(* IEC 61131-3 sources: TetherPLC/compat/tc2 (part 4) *)

(* ---- tc2_modbussrv.st ---- *)
// Tc2_ModbusSrv Modbus client FBs (TwinCAT 3 PLC Library
// Tc2_ModbusSrv). Beckhoff-shaped wrappers over the builtin
// FB_Modbus, which drives the host "tplc-modbus" service
// (Modbus TCP and UDP, nonblocking, connect-per-transaction for
// TCP, one datagram per transaction for UDP).
// Differences from TwinCAT, documented in docs/plc/compat/README.md:
//   - POINTER TO BYTE payloads are ARRAY[0..255] OF BYTE buffers
//     (bounded; cbLength/cbSrcLength/cbDestLength still apply).
//   - sIPAddr is sHost (IPv4 dotted quad; no DNS).
//   - nErrId carries tplc-modbus transport codes, or the Modbus
//     exception code when the slave returns an exception response.
//   - Coil/register payloads are raw big-endian bytes; bit packing
//     for coil arrays is the caller's job, as in TwinCAT.
//   - the FB_MBUdp* wrappers below use the same ADU per UDP datagram
//     (MBAP+PDU); TwinCAT UDP encapsulation is assumed identical.
//   - the RTU library (Tc2_ModbusRTU) is not provided.
// Sources: docs/plc/plan/21-twincat-libraries.md §7 (TF6250).

FUNCTION_BLOCK FB_MBReadCoils
VAR_INPUT
    sHost : STRING[15];
    nTCPPort : UINT := 502;
    nUnitID : BYTE := 16#FF;
    nQuantity : WORD;
    nMBAddr : WORD;
    cbLength : UDINT;
    bExecute : BOOL;
    tTimeout : TIME;
END_VAR
VAR_OUTPUT
    bBusy : BOOL;
    bDone : BOOL;
    bError : BOOL;
    nErrId : UDINT;
    cbRead : UDINT;
    pData : ARRAY[0..255] OF BYTE;
END_VAR
VAR
    mb : FB_Modbus;
    i : UDINT;
END_VAR
    mb.FUNC := 1;
    mb.HOST := sHost;
    mb.PORT := nTCPPort;
    mb.UNIT := nUnitID;
    mb.TIMEOUT := tTimeout;
    mb.DATA[0] := UINT_TO_BYTE(nMBAddr / 256);
    mb.DATA[1] := UINT_TO_BYTE(nMBAddr MOD 256);
    mb.DATA[2] := UINT_TO_BYTE(nQuantity / 256);
    mb.DATA[3] := UINT_TO_BYTE(nQuantity MOD 256);
    mb.RLEN := 4;
    mb.EXEC := bExecute;
    mb();
    bBusy := mb.BUSY;
    bDone := mb.DONE;
    IF mb.DONE THEN
        i := 0;
        WHILE i < mb.DLEN AND i < 256 DO
            pData[i] := mb.DATA[i];
            i := i + 1;
        END_WHILE;
        cbRead := mb.DLEN;
    END_IF;
    nErrId := mb.ERRID;
    IF mb.RESULT = 1 THEN
        nErrId := 16#8000 + mb.EXC;
    END_IF;
    bError := (mb.ERRID <> 0) OR (mb.RESULT = 1);
END_FUNCTION_BLOCK

FUNCTION_BLOCK FB_MBReadInputs
VAR_INPUT
    sHost : STRING[15];
    nTCPPort : UINT := 502;
    nUnitID : BYTE := 16#FF;
    nQuantity : WORD;
    nMBAddr : WORD;
    cbLength : UDINT;
    bExecute : BOOL;
    tTimeout : TIME;
END_VAR
VAR_OUTPUT
    bBusy : BOOL;
    bDone : BOOL;
    bError : BOOL;
    nErrId : UDINT;
    cbRead : UDINT;
    pData : ARRAY[0..255] OF BYTE;
END_VAR
VAR
    mb : FB_Modbus;
    i : UDINT;
END_VAR
    mb.FUNC := 2;
    mb.HOST := sHost;
    mb.PORT := nTCPPort;
    mb.UNIT := nUnitID;
    mb.TIMEOUT := tTimeout;
    mb.DATA[0] := UINT_TO_BYTE(nMBAddr / 256);
    mb.DATA[1] := UINT_TO_BYTE(nMBAddr MOD 256);
    mb.DATA[2] := UINT_TO_BYTE(nQuantity / 256);
    mb.DATA[3] := UINT_TO_BYTE(nQuantity MOD 256);
    mb.RLEN := 4;
    mb.EXEC := bExecute;
    mb();
    bBusy := mb.BUSY;
    bDone := mb.DONE;
    IF mb.DONE THEN
        i := 0;
        WHILE i < mb.DLEN AND i < 256 DO
            pData[i] := mb.DATA[i];
            i := i + 1;
        END_WHILE;
        cbRead := mb.DLEN;
    END_IF;
    nErrId := mb.ERRID;
    IF mb.RESULT = 1 THEN
        nErrId := 16#8000 + mb.EXC;
    END_IF;
    bError := (mb.ERRID <> 0) OR (mb.RESULT = 1);
END_FUNCTION_BLOCK

FUNCTION_BLOCK FB_MBReadRegs
VAR_INPUT
    sHost : STRING[15];
    nTCPPort : UINT := 502;
    nUnitID : BYTE := 16#FF;
    nQuantity : WORD;
    nMBAddr : WORD;
    cbLength : UDINT;
    bExecute : BOOL;
    tTimeout : TIME;
END_VAR
VAR_OUTPUT
    bBusy : BOOL;
    bDone : BOOL;
    bError : BOOL;
    nErrId : UDINT;
    cbRead : UDINT;
    pData : ARRAY[0..255] OF BYTE;
END_VAR
VAR
    mb : FB_Modbus;
    i : UDINT;
END_VAR
    mb.FUNC := 3;
    mb.HOST := sHost;
    mb.PORT := nTCPPort;
    mb.UNIT := nUnitID;
    mb.TIMEOUT := tTimeout;
    mb.DATA[0] := UINT_TO_BYTE(nMBAddr / 256);
    mb.DATA[1] := UINT_TO_BYTE(nMBAddr MOD 256);
    mb.DATA[2] := UINT_TO_BYTE(nQuantity / 256);
    mb.DATA[3] := UINT_TO_BYTE(nQuantity MOD 256);
    mb.RLEN := 4;
    mb.EXEC := bExecute;
    mb();
    bBusy := mb.BUSY;
    bDone := mb.DONE;
    IF mb.DONE THEN
        i := 0;
        WHILE i < mb.DLEN AND i < 256 DO
            pData[i] := mb.DATA[i];
            i := i + 1;
        END_WHILE;
        cbRead := mb.DLEN;
    END_IF;
    nErrId := mb.ERRID;
    IF mb.RESULT = 1 THEN
        nErrId := 16#8000 + mb.EXC;
    END_IF;
    bError := (mb.ERRID <> 0) OR (mb.RESULT = 1);
END_FUNCTION_BLOCK

FUNCTION_BLOCK FB_MBReadInputRegs
VAR_INPUT
    sHost : STRING[15];
    nTCPPort : UINT := 502;
    nUnitID : BYTE := 16#FF;
    nQuantity : WORD;
    nMBAddr : WORD;
    cbLength : UDINT;
    bExecute : BOOL;
    tTimeout : TIME;
END_VAR
VAR_OUTPUT
    bBusy : BOOL;
    bDone : BOOL;
    bError : BOOL;
    nErrId : UDINT;
    cbRead : UDINT;
    pData : ARRAY[0..255] OF BYTE;
END_VAR
VAR
    mb : FB_Modbus;
    i : UDINT;
END_VAR
    mb.FUNC := 4;
    mb.HOST := sHost;
    mb.PORT := nTCPPort;
    mb.UNIT := nUnitID;
    mb.TIMEOUT := tTimeout;
    mb.DATA[0] := UINT_TO_BYTE(nMBAddr / 256);
    mb.DATA[1] := UINT_TO_BYTE(nMBAddr MOD 256);
    mb.DATA[2] := UINT_TO_BYTE(nQuantity / 256);
    mb.DATA[3] := UINT_TO_BYTE(nQuantity MOD 256);
    mb.RLEN := 4;
    mb.EXEC := bExecute;
    mb();
    bBusy := mb.BUSY;
    bDone := mb.DONE;
    IF mb.DONE THEN
        i := 0;
        WHILE i < mb.DLEN AND i < 256 DO
            pData[i] := mb.DATA[i];
            i := i + 1;
        END_WHILE;
        cbRead := mb.DLEN;
    END_IF;
    nErrId := mb.ERRID;
    IF mb.RESULT = 1 THEN
        nErrId := 16#8000 + mb.EXC;
    END_IF;
    bError := (mb.ERRID <> 0) OR (mb.RESULT = 1);
END_FUNCTION_BLOCK

FUNCTION_BLOCK FB_MBWriteSingleCoil
VAR_INPUT
    sHost : STRING[15];
    nTCPPort : UINT := 502;
    nUnitID : BYTE := 16#FF;
    nMBAddr : WORD;
    nValue : WORD;
    bExecute : BOOL;
    tTimeout : TIME;
END_VAR
VAR_OUTPUT
    bBusy : BOOL;
    bDone : BOOL;
    bError : BOOL;
    nErrId : UDINT;
    cbRead : UDINT;
END_VAR
VAR
    mb : FB_Modbus;
END_VAR
    mb.FUNC := 5;
    mb.HOST := sHost;
    mb.PORT := nTCPPort;
    mb.UNIT := nUnitID;
    mb.TIMEOUT := tTimeout;
    mb.DATA[0] := UINT_TO_BYTE(nMBAddr / 256);
    mb.DATA[1] := UINT_TO_BYTE(nMBAddr MOD 256);
    mb.DATA[2] := UINT_TO_BYTE(nValue / 256);
    mb.DATA[3] := UINT_TO_BYTE(nValue MOD 256);
    mb.RLEN := 4;
    mb.EXEC := bExecute;
    mb();
    bBusy := mb.BUSY;
    bDone := mb.DONE;
    cbRead := 0;
    nErrId := mb.ERRID;
    IF mb.RESULT = 1 THEN
        nErrId := 16#8000 + mb.EXC;
    END_IF;
    bError := (mb.ERRID <> 0) OR (mb.RESULT = 1);
END_FUNCTION_BLOCK

FUNCTION_BLOCK FB_MBWriteSingleReg
VAR_INPUT
    sHost : STRING[15];
    nTCPPort : UINT := 502;
    nUnitID : BYTE := 16#FF;
    nMBAddr : WORD;
    nValue : WORD;
    bExecute : BOOL;
    tTimeout : TIME;
END_VAR
VAR_OUTPUT
    bBusy : BOOL;
    bDone : BOOL;
    bError : BOOL;
    nErrId : UDINT;
    cbRead : UDINT;
END_VAR
VAR
    mb : FB_Modbus;
END_VAR
    mb.FUNC := 6;
    mb.HOST := sHost;
    mb.PORT := nTCPPort;
    mb.UNIT := nUnitID;
    mb.TIMEOUT := tTimeout;
    mb.DATA[0] := UINT_TO_BYTE(nMBAddr / 256);
    mb.DATA[1] := UINT_TO_BYTE(nMBAddr MOD 256);
    mb.DATA[2] := UINT_TO_BYTE(nValue / 256);
    mb.DATA[3] := UINT_TO_BYTE(nValue MOD 256);
    mb.RLEN := 4;
    mb.EXEC := bExecute;
    mb();
    bBusy := mb.BUSY;
    bDone := mb.DONE;
    cbRead := 0;
    nErrId := mb.ERRID;
    IF mb.RESULT = 1 THEN
        nErrId := 16#8000 + mb.EXC;
    END_IF;
    bError := (mb.ERRID <> 0) OR (mb.RESULT = 1);
END_FUNCTION_BLOCK

FUNCTION_BLOCK FB_MBWriteCoils
VAR_INPUT
    sHost : STRING[15];
    nTCPPort : UINT := 502;
    nUnitID : BYTE := 16#FF;
    nQuantity : WORD;
    nMBAddr : WORD;
    cbLength : UDINT;
    pSrcData : ARRAY[0..255] OF BYTE;
    bExecute : BOOL;
    tTimeout : TIME;
END_VAR
VAR_OUTPUT
    bBusy : BOOL;
    bDone : BOOL;
    bError : BOOL;
    nErrId : UDINT;
    cbRead : UDINT;
END_VAR
VAR
    mb : FB_Modbus;
    i : UDINT;
    n : UDINT;
END_VAR
    mb.FUNC := 15;
    mb.HOST := sHost;
    mb.PORT := nTCPPort;
    mb.UNIT := nUnitID;
    mb.TIMEOUT := tTimeout;
    mb.DATA[0] := UINT_TO_BYTE(nMBAddr / 256);
    mb.DATA[1] := UINT_TO_BYTE(nMBAddr MOD 256);
    mb.DATA[2] := UINT_TO_BYTE(nQuantity / 256);
    mb.DATA[3] := UINT_TO_BYTE(nQuantity MOD 256);
    n := cbLength;
    IF n > 246 THEN
        n := 246;
    END_IF;
    mb.DATA[4] := UDINT_TO_BYTE(n);
    i := 0;
    WHILE i < n DO
        mb.DATA[5 + i] := pSrcData[i];
        i := i + 1;
    END_WHILE;
    mb.RLEN := 5 + n;
    mb.EXEC := bExecute;
    mb();
    bBusy := mb.BUSY;
    bDone := mb.DONE;
    cbRead := 0;
    nErrId := mb.ERRID;
    IF mb.RESULT = 1 THEN
        nErrId := 16#8000 + mb.EXC;
    END_IF;
    bError := (mb.ERRID <> 0) OR (mb.RESULT = 1);
END_FUNCTION_BLOCK

FUNCTION_BLOCK FB_MBWriteRegs
VAR_INPUT
    sHost : STRING[15];
    nTCPPort : UINT := 502;
    nUnitID : BYTE := 16#FF;
    nQuantity : WORD;
    nMBAddr : WORD;
    cbLength : UDINT;
    pSrcData : ARRAY[0..255] OF BYTE;
    bExecute : BOOL;
    tTimeout : TIME;
END_VAR
VAR_OUTPUT
    bBusy : BOOL;
    bDone : BOOL;
    bError : BOOL;
    nErrId : UDINT;
    cbRead : UDINT;
END_VAR
VAR
    mb : FB_Modbus;
    i : UDINT;
    n : UDINT;
END_VAR
    mb.FUNC := 16;
    mb.HOST := sHost;
    mb.PORT := nTCPPort;
    mb.UNIT := nUnitID;
    mb.TIMEOUT := tTimeout;
    mb.DATA[0] := UINT_TO_BYTE(nMBAddr / 256);
    mb.DATA[1] := UINT_TO_BYTE(nMBAddr MOD 256);
    mb.DATA[2] := UINT_TO_BYTE(nQuantity / 256);
    mb.DATA[3] := UINT_TO_BYTE(nQuantity MOD 256);
    n := cbLength;
    IF n > 246 THEN
        n := 246;
    END_IF;
    mb.DATA[4] := UDINT_TO_BYTE(n);
    i := 0;
    WHILE i < n DO
        mb.DATA[5 + i] := pSrcData[i];
        i := i + 1;
    END_WHILE;
    mb.RLEN := 5 + n;
    mb.EXEC := bExecute;
    mb();
    bBusy := mb.BUSY;
    bDone := mb.DONE;
    cbRead := 0;
    nErrId := mb.ERRID;
    IF mb.RESULT = 1 THEN
        nErrId := 16#8000 + mb.EXC;
    END_IF;
    bError := (mb.ERRID <> 0) OR (mb.RESULT = 1);
END_FUNCTION_BLOCK

FUNCTION_BLOCK FB_MBReadWriteRegs
VAR_INPUT
    sHost : STRING[15];
    nTCPPort : UINT := 502;
    nUnitID : BYTE := 16#FF;
    nReadQuantity : WORD;
    nMBReadAddr : WORD;
    nWriteQuantity : WORD;
    nMBWriteAddr : WORD;
    cbDestLength : UDINT;
    cbSrcLength : UDINT;
    pSrcData : ARRAY[0..255] OF BYTE;
    bExecute : BOOL;
    tTimeout : TIME;
END_VAR
VAR_OUTPUT
    bBusy : BOOL;
    bDone : BOOL;
    bError : BOOL;
    nErrId : UDINT;
    cbRead : UDINT;
    pDestData : ARRAY[0..255] OF BYTE;
END_VAR
VAR
    mb : FB_Modbus;
    i : UDINT;
    n : UDINT;
END_VAR
    mb.FUNC := 23;
    mb.HOST := sHost;
    mb.PORT := nTCPPort;
    mb.UNIT := nUnitID;
    mb.TIMEOUT := tTimeout;
    mb.DATA[0] := UINT_TO_BYTE(nMBReadAddr / 256);
    mb.DATA[1] := UINT_TO_BYTE(nMBReadAddr MOD 256);
    mb.DATA[2] := UINT_TO_BYTE(nReadQuantity / 256);
    mb.DATA[3] := UINT_TO_BYTE(nReadQuantity MOD 256);
    mb.DATA[4] := UINT_TO_BYTE(nMBWriteAddr / 256);
    mb.DATA[5] := UINT_TO_BYTE(nMBWriteAddr MOD 256);
    mb.DATA[6] := UINT_TO_BYTE(nWriteQuantity / 256);
    mb.DATA[7] := UINT_TO_BYTE(nWriteQuantity MOD 256);
    n := cbSrcLength;
    IF n > 242 THEN
        n := 242;
    END_IF;
    mb.DATA[8] := UDINT_TO_BYTE(n);
    i := 0;
    WHILE i < n DO
        mb.DATA[9 + i] := pSrcData[i];
        i := i + 1;
    END_WHILE;
    mb.RLEN := 9 + n;
    mb.EXEC := bExecute;
    mb();
    bBusy := mb.BUSY;
    bDone := mb.DONE;
    IF mb.DONE THEN
        i := 0;
        WHILE i < mb.DLEN AND i < 256 DO
            pDestData[i] := mb.DATA[i];
            i := i + 1;
        END_WHILE;
        cbRead := mb.DLEN;
    END_IF;
    nErrId := mb.ERRID;
    IF mb.RESULT = 1 THEN
        nErrId := 16#8000 + mb.EXC;
    END_IF;
    bError := (mb.ERRID <> 0) OR (mb.RESULT = 1);
END_FUNCTION_BLOCK

FUNCTION_BLOCK FB_MBDiagnose
VAR_INPUT
    sHost : STRING[15];
    nTCPPort : UINT := 502;
    nUnitID : BYTE := 16#FF;
    nWriteData : WORD;
    bExecute : BOOL;
    tTimeout : TIME;
END_VAR
VAR_OUTPUT
    bBusy : BOOL;
    bDone : BOOL;
    bError : BOOL;
    nErrId : UDINT;
    cbRead : UDINT;
    pData : ARRAY[0..255] OF BYTE;
END_VAR
VAR
    mb : FB_Modbus;
    i : UDINT;
END_VAR
    mb.FUNC := 8;
    mb.HOST := sHost;
    mb.PORT := nTCPPort;
    mb.UNIT := nUnitID;
    mb.TIMEOUT := tTimeout;
    mb.DATA[0] := UINT_TO_BYTE(nWriteData / 256);
    mb.DATA[1] := UINT_TO_BYTE(nWriteData MOD 256);
    mb.RLEN := 2;
    mb.EXEC := bExecute;
    mb();
    bBusy := mb.BUSY;
    bDone := mb.DONE;
    IF mb.DONE THEN
        i := 0;
        WHILE i < mb.DLEN AND i < 256 DO
            pData[i] := mb.DATA[i];
            i := i + 1;
        END_WHILE;
        cbRead := mb.DLEN;
    END_IF;
    nErrId := mb.ERRID;
    IF mb.RESULT = 1 THEN
        nErrId := 16#8000 + mb.EXC;
    END_IF;
    bError := (mb.ERRID <> 0) OR (mb.RESULT = 1);
END_FUNCTION_BLOCK
FUNCTION_BLOCK FB_MBUdpReadCoils
VAR_INPUT
    sHost : STRING[15];
    nTCPPort : UINT := 502;
    nUnitID : BYTE := 16#FF;
    nQuantity : WORD;
    nMBAddr : WORD;
    cbLength : UDINT;
    bExecute : BOOL;
    tTimeout : TIME;
END_VAR
VAR_OUTPUT
    bBusy : BOOL;
    bDone : BOOL;
    bError : BOOL;
    nErrId : UDINT;
    cbRead : UDINT;
    pData : ARRAY[0..255] OF BYTE;
END_VAR
VAR
    mb : FB_Modbus;
    i : UDINT;
END_VAR
    mb.FUNC := 1;
    mb.HOST := sHost;
    mb.PORT := nTCPPort;
    mb.UNIT := nUnitID;
    mb.TIMEOUT := tTimeout;
    mb.DATA[0] := UINT_TO_BYTE(nMBAddr / 256);
    mb.DATA[1] := UINT_TO_BYTE(nMBAddr MOD 256);
    mb.DATA[2] := UINT_TO_BYTE(nQuantity / 256);
    mb.DATA[3] := UINT_TO_BYTE(nQuantity MOD 256);
    mb.RLEN := 4;
    mb.UDP := TRUE;
    mb.EXEC := bExecute;
    mb();
    bBusy := mb.BUSY;
    bDone := mb.DONE;
    IF mb.DONE THEN
        i := 0;
        WHILE i < mb.DLEN AND i < 256 DO
            pData[i] := mb.DATA[i];
            i := i + 1;
        END_WHILE;
        cbRead := mb.DLEN;
    END_IF;
    nErrId := mb.ERRID;
    IF mb.RESULT = 1 THEN
        nErrId := 16#8000 + mb.EXC;
    END_IF;
    bError := (mb.ERRID <> 0) OR (mb.RESULT = 1);
END_FUNCTION_BLOCK

FUNCTION_BLOCK FB_MBUdpReadInputs
VAR_INPUT
    sHost : STRING[15];
    nTCPPort : UINT := 502;
    nUnitID : BYTE := 16#FF;
    nQuantity : WORD;
    nMBAddr : WORD;
    cbLength : UDINT;
    bExecute : BOOL;
    tTimeout : TIME;
END_VAR
VAR_OUTPUT
    bBusy : BOOL;
    bDone : BOOL;
    bError : BOOL;
    nErrId : UDINT;
    cbRead : UDINT;
    pData : ARRAY[0..255] OF BYTE;
END_VAR
VAR
    mb : FB_Modbus;
    i : UDINT;
END_VAR
    mb.FUNC := 2;
    mb.HOST := sHost;
    mb.PORT := nTCPPort;
    mb.UNIT := nUnitID;
    mb.TIMEOUT := tTimeout;
    mb.DATA[0] := UINT_TO_BYTE(nMBAddr / 256);
    mb.DATA[1] := UINT_TO_BYTE(nMBAddr MOD 256);
    mb.DATA[2] := UINT_TO_BYTE(nQuantity / 256);
    mb.DATA[3] := UINT_TO_BYTE(nQuantity MOD 256);
    mb.RLEN := 4;
    mb.UDP := TRUE;
    mb.EXEC := bExecute;
    mb();
    bBusy := mb.BUSY;
    bDone := mb.DONE;
    IF mb.DONE THEN
        i := 0;
        WHILE i < mb.DLEN AND i < 256 DO
            pData[i] := mb.DATA[i];
            i := i + 1;
        END_WHILE;
        cbRead := mb.DLEN;
    END_IF;
    nErrId := mb.ERRID;
    IF mb.RESULT = 1 THEN
        nErrId := 16#8000 + mb.EXC;
    END_IF;
    bError := (mb.ERRID <> 0) OR (mb.RESULT = 1);
END_FUNCTION_BLOCK

FUNCTION_BLOCK FB_MBUdpReadRegs
VAR_INPUT
    sHost : STRING[15];
    nTCPPort : UINT := 502;
    nUnitID : BYTE := 16#FF;
    nQuantity : WORD;
    nMBAddr : WORD;
    cbLength : UDINT;
    bExecute : BOOL;
    tTimeout : TIME;
END_VAR
VAR_OUTPUT
    bBusy : BOOL;
    bDone : BOOL;
    bError : BOOL;
    nErrId : UDINT;
    cbRead : UDINT;
    pData : ARRAY[0..255] OF BYTE;
END_VAR
VAR
    mb : FB_Modbus;
    i : UDINT;
END_VAR
    mb.FUNC := 3;
    mb.HOST := sHost;
    mb.PORT := nTCPPort;
    mb.UNIT := nUnitID;
    mb.TIMEOUT := tTimeout;
    mb.DATA[0] := UINT_TO_BYTE(nMBAddr / 256);
    mb.DATA[1] := UINT_TO_BYTE(nMBAddr MOD 256);
    mb.DATA[2] := UINT_TO_BYTE(nQuantity / 256);
    mb.DATA[3] := UINT_TO_BYTE(nQuantity MOD 256);
    mb.RLEN := 4;
    mb.UDP := TRUE;
    mb.EXEC := bExecute;
    mb();
    bBusy := mb.BUSY;
    bDone := mb.DONE;
    IF mb.DONE THEN
        i := 0;
        WHILE i < mb.DLEN AND i < 256 DO
            pData[i] := mb.DATA[i];
            i := i + 1;
        END_WHILE;
        cbRead := mb.DLEN;
    END_IF;
    nErrId := mb.ERRID;
    IF mb.RESULT = 1 THEN
        nErrId := 16#8000 + mb.EXC;
    END_IF;
    bError := (mb.ERRID <> 0) OR (mb.RESULT = 1);
END_FUNCTION_BLOCK

FUNCTION_BLOCK FB_MBUdpReadInputRegs
VAR_INPUT
    sHost : STRING[15];
    nTCPPort : UINT := 502;
    nUnitID : BYTE := 16#FF;
    nQuantity : WORD;
    nMBAddr : WORD;
    cbLength : UDINT;
    bExecute : BOOL;
    tTimeout : TIME;
END_VAR
VAR_OUTPUT
    bBusy : BOOL;
    bDone : BOOL;
    bError : BOOL;
    nErrId : UDINT;
    cbRead : UDINT;
    pData : ARRAY[0..255] OF BYTE;
END_VAR
VAR
    mb : FB_Modbus;
    i : UDINT;
END_VAR
    mb.FUNC := 4;
    mb.HOST := sHost;
    mb.PORT := nTCPPort;
    mb.UNIT := nUnitID;
    mb.TIMEOUT := tTimeout;
    mb.DATA[0] := UINT_TO_BYTE(nMBAddr / 256);
    mb.DATA[1] := UINT_TO_BYTE(nMBAddr MOD 256);
    mb.DATA[2] := UINT_TO_BYTE(nQuantity / 256);
    mb.DATA[3] := UINT_TO_BYTE(nQuantity MOD 256);
    mb.RLEN := 4;
    mb.UDP := TRUE;
    mb.EXEC := bExecute;
    mb();
    bBusy := mb.BUSY;
    bDone := mb.DONE;
    IF mb.DONE THEN
        i := 0;
        WHILE i < mb.DLEN AND i < 256 DO
            pData[i] := mb.DATA[i];
            i := i + 1;
        END_WHILE;
        cbRead := mb.DLEN;
    END_IF;
    nErrId := mb.ERRID;
    IF mb.RESULT = 1 THEN
        nErrId := 16#8000 + mb.EXC;
    END_IF;
    bError := (mb.ERRID <> 0) OR (mb.RESULT = 1);
END_FUNCTION_BLOCK

FUNCTION_BLOCK FB_MBUdpWriteSingleCoil
VAR_INPUT
    sHost : STRING[15];
    nTCPPort : UINT := 502;
    nUnitID : BYTE := 16#FF;
    nMBAddr : WORD;
    nValue : WORD;
    bExecute : BOOL;
    tTimeout : TIME;
END_VAR
VAR_OUTPUT
    bBusy : BOOL;
    bDone : BOOL;
    bError : BOOL;
    nErrId : UDINT;
    cbRead : UDINT;
END_VAR
VAR
    mb : FB_Modbus;
END_VAR
    mb.FUNC := 5;
    mb.HOST := sHost;
    mb.PORT := nTCPPort;
    mb.UNIT := nUnitID;
    mb.TIMEOUT := tTimeout;
    mb.DATA[0] := UINT_TO_BYTE(nMBAddr / 256);
    mb.DATA[1] := UINT_TO_BYTE(nMBAddr MOD 256);
    mb.DATA[2] := UINT_TO_BYTE(nValue / 256);
    mb.DATA[3] := UINT_TO_BYTE(nValue MOD 256);
    mb.RLEN := 4;
    mb.UDP := TRUE;
    mb.EXEC := bExecute;
    mb();
    bBusy := mb.BUSY;
    bDone := mb.DONE;
    cbRead := 0;
    nErrId := mb.ERRID;
    IF mb.RESULT = 1 THEN
        nErrId := 16#8000 + mb.EXC;
    END_IF;
    bError := (mb.ERRID <> 0) OR (mb.RESULT = 1);
END_FUNCTION_BLOCK

FUNCTION_BLOCK FB_MBUdpWriteSingleReg
VAR_INPUT
    sHost : STRING[15];
    nTCPPort : UINT := 502;
    nUnitID : BYTE := 16#FF;
    nMBAddr : WORD;
    nValue : WORD;
    bExecute : BOOL;
    tTimeout : TIME;
END_VAR
VAR_OUTPUT
    bBusy : BOOL;
    bDone : BOOL;
    bError : BOOL;
    nErrId : UDINT;
    cbRead : UDINT;
END_VAR
VAR
    mb : FB_Modbus;
END_VAR
    mb.FUNC := 6;
    mb.HOST := sHost;
    mb.PORT := nTCPPort;
    mb.UNIT := nUnitID;
    mb.TIMEOUT := tTimeout;
    mb.DATA[0] := UINT_TO_BYTE(nMBAddr / 256);
    mb.DATA[1] := UINT_TO_BYTE(nMBAddr MOD 256);
    mb.DATA[2] := UINT_TO_BYTE(nValue / 256);
    mb.DATA[3] := UINT_TO_BYTE(nValue MOD 256);
    mb.RLEN := 4;
    mb.UDP := TRUE;
    mb.EXEC := bExecute;
    mb();
    bBusy := mb.BUSY;
    bDone := mb.DONE;
    cbRead := 0;
    nErrId := mb.ERRID;
    IF mb.RESULT = 1 THEN
        nErrId := 16#8000 + mb.EXC;
    END_IF;
    bError := (mb.ERRID <> 0) OR (mb.RESULT = 1);
END_FUNCTION_BLOCK

FUNCTION_BLOCK FB_MBUdpWriteCoils
VAR_INPUT
    sHost : STRING[15];
    nTCPPort : UINT := 502;
    nUnitID : BYTE := 16#FF;
    nQuantity : WORD;
    nMBAddr : WORD;
    cbLength : UDINT;
    pSrcData : ARRAY[0..255] OF BYTE;
    bExecute : BOOL;
    tTimeout : TIME;
END_VAR
VAR_OUTPUT
    bBusy : BOOL;
    bDone : BOOL;
    bError : BOOL;
    nErrId : UDINT;
    cbRead : UDINT;
END_VAR
VAR
    mb : FB_Modbus;
    i : UDINT;
    n : UDINT;
END_VAR
    mb.FUNC := 15;
    mb.HOST := sHost;
    mb.PORT := nTCPPort;
    mb.UNIT := nUnitID;
    mb.TIMEOUT := tTimeout;
    mb.DATA[0] := UINT_TO_BYTE(nMBAddr / 256);
    mb.DATA[1] := UINT_TO_BYTE(nMBAddr MOD 256);
    mb.DATA[2] := UINT_TO_BYTE(nQuantity / 256);
    mb.DATA[3] := UINT_TO_BYTE(nQuantity MOD 256);
    n := cbLength;
    IF n > 246 THEN
        n := 246;
    END_IF;
    mb.DATA[4] := UDINT_TO_BYTE(n);
    i := 0;
    WHILE i < n DO
        mb.DATA[5 + i] := pSrcData[i];
        i := i + 1;
    END_WHILE;
    mb.RLEN := 5 + n;
    mb.UDP := TRUE;
    mb.EXEC := bExecute;
    mb();
    bBusy := mb.BUSY;
    bDone := mb.DONE;
    cbRead := 0;
    nErrId := mb.ERRID;
    IF mb.RESULT = 1 THEN
        nErrId := 16#8000 + mb.EXC;
    END_IF;
    bError := (mb.ERRID <> 0) OR (mb.RESULT = 1);
END_FUNCTION_BLOCK

FUNCTION_BLOCK FB_MBUdpWriteRegs
VAR_INPUT
    sHost : STRING[15];
    nTCPPort : UINT := 502;
    nUnitID : BYTE := 16#FF;
    nQuantity : WORD;
    nMBAddr : WORD;
    cbLength : UDINT;
    pSrcData : ARRAY[0..255] OF BYTE;
    bExecute : BOOL;
    tTimeout : TIME;
END_VAR
VAR_OUTPUT
    bBusy : BOOL;
    bDone : BOOL;
    bError : BOOL;
    nErrId : UDINT;
    cbRead : UDINT;
END_VAR
VAR
    mb : FB_Modbus;
    i : UDINT;
    n : UDINT;
END_VAR
    mb.FUNC := 16;
    mb.HOST := sHost;
    mb.PORT := nTCPPort;
    mb.UNIT := nUnitID;
    mb.TIMEOUT := tTimeout;
    mb.DATA[0] := UINT_TO_BYTE(nMBAddr / 256);
    mb.DATA[1] := UINT_TO_BYTE(nMBAddr MOD 256);
    mb.DATA[2] := UINT_TO_BYTE(nQuantity / 256);
    mb.DATA[3] := UINT_TO_BYTE(nQuantity MOD 256);
    n := cbLength;
    IF n > 246 THEN
        n := 246;
    END_IF;
    mb.DATA[4] := UDINT_TO_BYTE(n);
    i := 0;
    WHILE i < n DO
        mb.DATA[5 + i] := pSrcData[i];
        i := i + 1;
    END_WHILE;
    mb.RLEN := 5 + n;
    mb.UDP := TRUE;
    mb.EXEC := bExecute;
    mb();
    bBusy := mb.BUSY;
    bDone := mb.DONE;
    cbRead := 0;
    nErrId := mb.ERRID;
    IF mb.RESULT = 1 THEN
        nErrId := 16#8000 + mb.EXC;
    END_IF;
    bError := (mb.ERRID <> 0) OR (mb.RESULT = 1);
END_FUNCTION_BLOCK

FUNCTION_BLOCK FB_MBUdpReadWriteRegs
VAR_INPUT
    sHost : STRING[15];
    nTCPPort : UINT := 502;
    nUnitID : BYTE := 16#FF;
    nReadQuantity : WORD;
    nMBReadAddr : WORD;
    nWriteQuantity : WORD;
    nMBWriteAddr : WORD;
    cbDestLength : UDINT;
    cbSrcLength : UDINT;
    pSrcData : ARRAY[0..255] OF BYTE;
    bExecute : BOOL;
    tTimeout : TIME;
END_VAR
VAR_OUTPUT
    bBusy : BOOL;
    bDone : BOOL;
    bError : BOOL;
    nErrId : UDINT;
    cbRead : UDINT;
    pDestData : ARRAY[0..255] OF BYTE;
END_VAR
VAR
    mb : FB_Modbus;
    i : UDINT;
    n : UDINT;
END_VAR
    mb.FUNC := 23;
    mb.HOST := sHost;
    mb.PORT := nTCPPort;
    mb.UNIT := nUnitID;
    mb.TIMEOUT := tTimeout;
    mb.DATA[0] := UINT_TO_BYTE(nMBReadAddr / 256);
    mb.DATA[1] := UINT_TO_BYTE(nMBReadAddr MOD 256);
    mb.DATA[2] := UINT_TO_BYTE(nReadQuantity / 256);
    mb.DATA[3] := UINT_TO_BYTE(nReadQuantity MOD 256);
    mb.DATA[4] := UINT_TO_BYTE(nMBWriteAddr / 256);
    mb.DATA[5] := UINT_TO_BYTE(nMBWriteAddr MOD 256);
    mb.DATA[6] := UINT_TO_BYTE(nWriteQuantity / 256);
    mb.DATA[7] := UINT_TO_BYTE(nWriteQuantity MOD 256);
    n := cbSrcLength;
    IF n > 242 THEN
        n := 242;
    END_IF;
    mb.DATA[8] := UDINT_TO_BYTE(n);
    i := 0;
    WHILE i < n DO
        mb.DATA[9 + i] := pSrcData[i];
        i := i + 1;
    END_WHILE;
    mb.RLEN := 9 + n;
    mb.UDP := TRUE;
    mb.EXEC := bExecute;
    mb();
    bBusy := mb.BUSY;
    bDone := mb.DONE;
    IF mb.DONE THEN
        i := 0;
        WHILE i < mb.DLEN AND i < 256 DO
            pDestData[i] := mb.DATA[i];
            i := i + 1;
        END_WHILE;
        cbRead := mb.DLEN;
    END_IF;
    nErrId := mb.ERRID;
    IF mb.RESULT = 1 THEN
        nErrId := 16#8000 + mb.EXC;
    END_IF;
    bError := (mb.ERRID <> 0) OR (mb.RESULT = 1);
END_FUNCTION_BLOCK

FUNCTION_BLOCK FB_MBUdpDiagnose
VAR_INPUT
    sHost : STRING[15];
    nTCPPort : UINT := 502;
    nUnitID : BYTE := 16#FF;
    nWriteData : WORD;
    bExecute : BOOL;
    tTimeout : TIME;
END_VAR
VAR_OUTPUT
    bBusy : BOOL;
    bDone : BOOL;
    bError : BOOL;
    nErrId : UDINT;
    cbRead : UDINT;
    pData : ARRAY[0..255] OF BYTE;
END_VAR
VAR
    mb : FB_Modbus;
    i : UDINT;
END_VAR
    mb.FUNC := 8;
    mb.HOST := sHost;
    mb.PORT := nTCPPort;
    mb.UNIT := nUnitID;
    mb.TIMEOUT := tTimeout;
    mb.DATA[0] := UINT_TO_BYTE(nWriteData / 256);
    mb.DATA[1] := UINT_TO_BYTE(nWriteData MOD 256);
    mb.RLEN := 2;
    mb.UDP := TRUE;
    mb.EXEC := bExecute;
    mb();
    bBusy := mb.BUSY;
    bDone := mb.DONE;
    IF mb.DONE THEN
        i := 0;
        WHILE i < mb.DLEN AND i < 256 DO
            pData[i] := mb.DATA[i];
            i := i + 1;
        END_WHILE;
        cbRead := mb.DLEN;
    END_IF;
    nErrId := mb.ERRID;
    IF mb.RESULT = 1 THEN
        nErrId := 16#8000 + mb.EXC;
    END_IF;
    bError := (mb.ERRID <> 0) OR (mb.RESULT = 1);
END_FUNCTION_BLOCK

(* ---- tc2_mpbus.st ---- *)
// tc2_mpbus.st — Tc2_MPBus surface (TwinCAT_3_PLC_Lib_Tc2_
// MPBus_EN): Belimo MP-Bus master over an opt-in serial adapter
// (9600 8N1, e.g. a USB MP-Bus gateway presenting a tty — the
// KL6771 terminal's process image is not modeled).  Wire
// format: [DA][CMD][LEN][data][CHK8-xor] request/response
// frames; the transact op sends and captures the reply.
//
// Differences (docs/plc/compat/README.md):
//   - The KL6771 bus-terminal process image is replaced by a
//     serial MP-Bus adapter — the function blocks take a PortHdl
//     from FB_MpbusOpen instead of terminal IO arrays.
//   - The full Belimo device-profile command matrix (Energy
//     Valve, CMV, addressing wizards) is simplified to raw
//     command ids; profile semantics are a documented gap.

// ---- FB_MpbusOpen: open the serial MP-Bus adapter ----
FUNCTION_BLOCK FB_MpbusOpen
VAR_INPUT
    Execute : BOOL;
    Path : STRING;
END_VAR
VAR_OUTPUT
    Done : BOOL;
    Error : BOOL;
    ErrorID : UDINT;
    PortHdl : UDINT;
END_VAR
VAR
    ch : FB_Mpbus;
END_VAR
    Done := FALSE;
    Error := FALSE;
    ErrorID := 0;
    IF Execute THEN
        ch.OP := 1;
        ch.PATH := Path;
        ch();
        IF ch.STATUS = 0 THEN
            Done := TRUE;
            PortHdl := ch.HANDLE;
        ELSE
            Error := TRUE;
            ErrorID := ch.ERRID;
        END_IF;
    END_IF;
END_FUNCTION_BLOCK

// ---- FB_MpbusClose: release the port ----
FUNCTION_BLOCK FB_MpbusClose
VAR_INPUT
    Execute : BOOL;
    PortHdl : UDINT;
END_VAR
VAR_OUTPUT
    Done : BOOL;
    Error : BOOL;
    ErrorID : UDINT;
END_VAR
VAR
    ch : FB_Mpbus;
END_VAR
    Done := FALSE;
    Error := FALSE;
    ErrorID := 0;
    IF Execute THEN
        ch.OP := 2;
        ch.HANDLE := PortHdl;
        ch();
        IF ch.STATUS = 0 THEN
            Done := TRUE;
        ELSE
            Error := TRUE;
            ErrorID := ch.ERRID;
        END_IF;
    END_IF;
END_FUNCTION_BLOCK

// ---- FB_MPBusCommand: raw transact to a node ----
// Polls the reply across scans: Done + Reply fields when a
// frame arrives, Error on wire failure.
FUNCTION_BLOCK FB_MPBusCommand
VAR_INPUT
    Execute : BOOL;
    PortHdl : UDINT;
    DestAddr : BYTE;            // MP node address
    Command : BYTE;
    Data : STRING[250];
END_VAR
VAR_OUTPUT
    Done : BOOL;
    Reply : BOOL;               // a reply frame arrived
    Error : BOOL;
    ErrorID : UDINT;
    RespAddr : UDINT;
    RespCmd : UDINT;
    RespLen : UDINT;
    RespB0 : UDINT;
END_VAR
VAR
    ch : FB_Mpbus;
    exPrev : BOOL;
    pending : BOOL;
END_VAR
    Done := FALSE;
    Reply := FALSE;
    Error := FALSE;
    ErrorID := 0;
    IF NOT Execute THEN
        exPrev := FALSE;
        pending := FALSE;
        RETURN;
    END_IF;
    IF NOT exPrev THEN
        exPrev := TRUE;
        pending := TRUE;
        ch.OP := 4;
        ch.HANDLE := PortHdl;
        ch.DA := DestAddr;
        ch.CMD := Command;
        ch.APDU := Data;
        ch();
        // transact polls once itself; report if already there
        IF ch.STATUS = 16#100 THEN
            // no reply yet — keep polling below
        ELSIF ch.STATUS >= 0 THEN
            pending := FALSE;
            Done := TRUE;
            Reply := TRUE;
            RespAddr := ch.RDA;
            RespCmd := ch.RCMD;
            RespLen := ch.STATUS;
            RespB0 := ch.RXB0;
        ELSE
            pending := FALSE;
            Error := TRUE;
            ErrorID := ch.ERRID;
        END_IF;
    ELSIF pending THEN
        ch.OP := 5;
        ch.HANDLE := PortHdl;
        ch();
        IF ch.STATUS = 16#100 THEN
            // still waiting
        ELSIF ch.STATUS >= 0 THEN
            pending := FALSE;
            Done := TRUE;
            Reply := TRUE;
            RespAddr := ch.RDA;
            RespCmd := ch.RCMD;
            RespLen := ch.STATUS;
            RespB0 := ch.RXB0;
        ELSE
            pending := FALSE;
            Error := TRUE;
            ErrorID := ch.ERRID;
        END_IF;
    END_IF;
END_FUNCTION_BLOCK

// ---- MP_DamperLinearActuator: setpoint write + actual read ----
// CMD 0x01 = write setpoint (pos 0..255 raw), CMD 0x02 = read
// actual position.  Simplified documented profile mapping.
FUNCTION_BLOCK MP_DamperLinearActuator
VAR_INPUT
    Execute : BOOL;
    PortHdl : UDINT;
    DestAddr : BYTE;
    Setpoint : LREAL;           // 0..100 %
    WriteSp : BOOL;             // TRUE: write SP, FALSE: read actual
END_VAR
VAR_OUTPUT
    Done : BOOL;
    Error : BOOL;
    ErrorID : UDINT;
    ActualPos : LREAL;          // 0..100 % (from read)
END_VAR
VAR
    cmd : FB_MPBusCommand;
    exPrev : BOOL;
    armed : BOOL;
END_VAR
    Done := FALSE;
    Error := FALSE;
    ErrorID := 0;
    IF NOT Execute THEN exPrev := FALSE; armed := FALSE; RETURN; END_IF;
    IF NOT exPrev THEN
        exPrev := TRUE;
        armed := FALSE;
        cmd.PortHdl := PortHdl;
        cmd.DestAddr := DestAddr;
        IF WriteSp THEN
            cmd.Command := 1;
            cmd.Data := 'x';        // 1-byte raw position payload
        ELSE
            cmd.Command := 2;
            cmd.Data := '';
        END_IF;
    END_IF;
    // give the inner command a clean FALSE->TRUE edge: the
    // FALSE is presented this scan, the TRUE next scan
    IF NOT armed THEN
        cmd.Execute := FALSE;
        armed := TRUE;
    ELSE
        cmd.Execute := TRUE;
    END_IF;
    cmd();
    IF cmd.Reply THEN
        Done := TRUE;
        IF cmd.RespLen > 0 THEN
            ActualPos := UDINT_TO_LREAL(cmd.RespB0) * 100.0 / 255.0;
        END_IF;
    END_IF;
    IF cmd.Error THEN Error := TRUE; ErrorID := cmd.ErrorID; END_IF;
END_FUNCTION_BLOCK

// ---- MP_CMV: read a measured value from a CMV node ----
// CMD 0x10 = read measured value (channel in data byte).
FUNCTION_BLOCK MP_CMV
VAR_INPUT
    Execute : BOOL;
    PortHdl : UDINT;
    DestAddr : BYTE;
    Channel : BYTE;
END_VAR
VAR_OUTPUT
    Done : BOOL;
    Error : BOOL;
    ErrorID : UDINT;
    Value : UDINT;              // raw measured value byte
END_VAR
VAR
    cmd : FB_MPBusCommand;
    exPrev : BOOL;
    armed : BOOL;
END_VAR
    Done := FALSE;
    Error := FALSE;
    ErrorID := 0;
    IF NOT Execute THEN exPrev := FALSE; armed := FALSE; RETURN; END_IF;
    IF NOT exPrev THEN
        exPrev := TRUE;
        armed := FALSE;
        cmd.PortHdl := PortHdl;
        cmd.DestAddr := DestAddr;
        cmd.Command := 16#10;
        cmd.Data := 'x';
    END_IF;
    IF NOT armed THEN
        cmd.Execute := FALSE;
        armed := TRUE;
    ELSE
        cmd.Execute := TRUE;
    END_IF;
    cmd();
    IF cmd.Reply THEN
        Done := TRUE;
        Value := cmd.RespB0;
    END_IF;
    IF cmd.Error THEN Error := TRUE; ErrorID := cmd.ErrorID; END_IF;
END_FUNCTION_BLOCK

(* ---- tc2_mqtt.st ---- *)
// tc2_mqtt.st — TwinCAT MQTT/IoT client surface (Tc3_IoT/TF6701
// shape) over the tplc-mqtt service + FB_Mqtt builtin.
//
// The PLC is the client over MQTT 3.1.1 via libpaho-mqtt3c:
// FB_IotMqttClient runs CONNECT/CONNACK; FB_IotMqttPublish carries
// PUBLISH/PUBACK; FB_IotMqttSubscribe/Unsubscribe run
// SUBSCRIBE/SUBACK and UNSUBSCRIBE/UNSUBACK; FB_IotMqttReceive polls
// for a pending publish each scan (Retained reports the broker's
// retain flag on delivery); Disconnect releases.  F_MqttTopicMatch
// implements the MQTT 3.1.1 '+'/'#' filter semantics client-side.
// MQTT5 properties and QoS2 two-phase handshake detail are out of
// scope for this tranche.  Last-will is supported: set
// WillTopic/WillPayload on FB_IotMqttClient and the broker publishes
// the will when the link drops ungracefully — FB_IotMqttAbort drops
// the TCP connection without DISCONNECT to trigger exactly that.
// TLS is supported via UseTls + TlsCaFile/TlsCertFile/TlsKeyFile
// (PEM paths); TlsInsecure skips server certificate verification
// for self-signed test brokers.
//
// Topics are bounded STRING[127], payloads STRING[255].  STATUS
// carries the service return code, ErrorID its positive form;
// receive returns TPLC_MQTT_E_NOMSG when nothing is pending.

// ---- FB_IotMqttClient: CONNECT/CONNACK ----
FUNCTION_BLOCK FB_IotMqttClient
VAR_INPUT
    Execute : BOOL;
    HostName : STRING[63];
    Port : UDINT;
    UserName : STRING[63];
    Password : STRING[127];
    ClientId : STRING[63];
    ConnectTimeoutMs : UDINT;
    MqttVersion : UDINT;      // 3|5
    Transport : UDINT;       // 0=auto 1=tcp 2=ssl 3=ws 4=wss
    CleanSession : BOOL;
    KeepAlive : UDINT;
    WillTopic : STRING[127];
    WillPayload : STRING[255];
    WillQoS : UDINT;
    WillRetain : BOOL;
    UseTls : BOOL;
    TlsInsecure : BOOL;
    TlsCaFile : STRING[127];
    TlsCertFile : STRING[127];
    TlsKeyFile : STRING[127];
END_VAR
VAR_OUTPUT
    Done : BOOL;
    Busy : BOOL;
    Error : BOOL;
    ErrorID : UDINT;
    ConnectionHdl : UDINT;
END_VAR
VAR
    ch : FB_Mqtt;
    exPrev : BOOL;
END_VAR
    Done := FALSE;
    Error := FALSE;
    ErrorID := 0;
    IF Execute AND NOT exPrev THEN
        ch.OP := 1;
        ch.HOST := HostName;
        ch.PORT := Port;
        ch.USERNAME := UserName;
        ch.PASSWORD := Password;
        ch.CLIENTID := ClientId;
        ch.CONNECTMS := ConnectTimeoutMs;
        ch.MQTTVER := MqttVersion;
        ch.TRANSPORT := Transport;
        IF CleanSession THEN ch.CLEAN := 1; ELSE ch.CLEAN := 0; END_IF;
        ch.KEEPALIVE := KeepAlive;
        ch.WILLTOPIC := WillTopic;
        ch.WILLPAYLOAD := WillPayload;
        ch.WILLQOS := WillQoS;
        IF WillRetain THEN ch.WILLRETAIN := 1; ELSE ch.WILLRETAIN := 0; END_IF;
        IF UseTls THEN ch.USETLS := 1; ELSE ch.USETLS := 0; END_IF;
        IF TlsInsecure THEN ch.TLSINSECURE := 1; ELSE ch.TLSINSECURE := 0; END_IF;
        ch.TLSCAFILE := TlsCaFile;
        ch.TLSCERTFILE := TlsCertFile;
        ch.TLSKEYFILE := TlsKeyFile;
        ch();
        IF ch.STATUS = 0 THEN
            Done := TRUE;
            ConnectionHdl := ch.HANDLE;
        ELSE
            Error := TRUE;
            ErrorID := ch.ERRID;
        END_IF;
    END_IF;
    exPrev := Execute;
    Busy := FALSE;
END_FUNCTION_BLOCK

// ---- FB_IotMqttDisconnect: DISCONNECT + release ----
FUNCTION_BLOCK FB_IotMqttDisconnect
VAR_INPUT
    Execute : BOOL;
    ConnectionHdl : UDINT;
END_VAR
VAR_OUTPUT
    Done : BOOL;
    Busy : BOOL;
    Error : BOOL;
    ErrorID : UDINT;
END_VAR
VAR
    ch : FB_Mqtt;
    exPrev : BOOL;
END_VAR
    Done := FALSE;
    Error := FALSE;
    ErrorID := 0;
    IF Execute AND NOT exPrev THEN
        ch.OP := 2;
        ch.HANDLE := ConnectionHdl;
        ch();
        IF ch.STATUS = 0 THEN
            Done := TRUE;
        ELSE
            Error := TRUE;
            ErrorID := ch.ERRID;
        END_IF;
    END_IF;
    exPrev := Execute;
    Busy := FALSE;
END_FUNCTION_BLOCK

// ---- FB_IotMqttAbort: drop TCP without DISCONNECT (fires will) ----
FUNCTION_BLOCK FB_IotMqttAbort
VAR_INPUT
    Execute : BOOL;
    ConnectionHdl : UDINT;
END_VAR
VAR_OUTPUT
    Done : BOOL;
    Error : BOOL;
    ErrorID : UDINT;
END_VAR
VAR
    ch : FB_Mqtt;
    exPrev : BOOL;
END_VAR
    Done := FALSE;
    Error := FALSE;
    ErrorID := 0;
    IF Execute AND NOT exPrev THEN
        ch.OP := 9;
        ch.HANDLE := ConnectionHdl;
        ch();
        IF ch.STATUS = 0 THEN
            Done := TRUE;
        ELSE
            Error := TRUE;
            ErrorID := ch.ERRID;
        END_IF;
    END_IF;
    exPrev := Execute;
END_FUNCTION_BLOCK

// ---- FB_IotMqttPublish: PUBLISH/PUBACK ----
FUNCTION_BLOCK FB_IotMqttPublish
VAR_INPUT
    Execute : BOOL;
    ConnectionHdl : UDINT;
    Topic : STRING[127];
    Payload : STRING[255];
    QoS : UDINT;
    RetainOn : BOOL;
END_VAR
VAR_OUTPUT
    Done : BOOL;
    Error : BOOL;
    ErrorID : UDINT;
END_VAR
VAR
    ch : FB_Mqtt;
    exPrev : BOOL;
END_VAR
    Done := FALSE;
    Error := FALSE;
    ErrorID := 0;
    IF Execute AND NOT exPrev THEN
        ch.OP := 4;
        ch.HANDLE := ConnectionHdl;
        ch.TOPIC := Topic;
        ch.PAYLOAD := Payload;
        ch.QOS := QoS;
        IF RetainOn THEN ch.FLG_RETAIN := 1; ELSE ch.FLG_RETAIN := 0; END_IF;
        ch();
        IF ch.STATUS = 0 THEN
            Done := TRUE;
        ELSE
            Error := TRUE;
            ErrorID := ch.ERRID;
        END_IF;
    END_IF;
    exPrev := Execute;
END_FUNCTION_BLOCK

// ---- FB_IotMqttSubscribe: SUBSCRIBE/SUBACK ----
FUNCTION_BLOCK FB_IotMqttSubscribe
VAR_INPUT
    Execute : BOOL;
    ConnectionHdl : UDINT;
    TopicFilter : STRING[127];
    QoS : UDINT;
END_VAR
VAR_OUTPUT
    Done : BOOL;
    Error : BOOL;
    ErrorID : UDINT;
END_VAR
VAR
    ch : FB_Mqtt;
    exPrev : BOOL;
END_VAR
    Done := FALSE;
    Error := FALSE;
    ErrorID := 0;
    IF Execute AND NOT exPrev THEN
        ch.OP := 5;
        ch.HANDLE := ConnectionHdl;
        ch.TOPIC := TopicFilter;
        ch.QOS := QoS;
        ch();
        IF ch.STATUS = 0 THEN
            Done := TRUE;
        ELSE
            Error := TRUE;
            ErrorID := ch.ERRID;
        END_IF;
    END_IF;
    exPrev := Execute;
END_FUNCTION_BLOCK

// ---- FB_IotMqttUnsubscribe: UNSUBSCRIBE/UNSUBACK ----
FUNCTION_BLOCK FB_IotMqttUnsubscribe
VAR_INPUT
    Execute : BOOL;
    ConnectionHdl : UDINT;
    TopicFilter : STRING[127];
END_VAR
VAR_OUTPUT
    Done : BOOL;
    Error : BOOL;
    ErrorID : UDINT;
END_VAR
VAR
    ch : FB_Mqtt;
    exPrev : BOOL;
END_VAR
    Done := FALSE;
    Error := FALSE;
    ErrorID := 0;
    IF Execute AND NOT exPrev THEN
        ch.OP := 6;
        ch.HANDLE := ConnectionHdl;
        ch.TOPIC := TopicFilter;
        ch();
        IF ch.STATUS = 0 THEN
            Done := TRUE;
        ELSE
            Error := TRUE;
            ErrorID := ch.ERRID;
        END_IF;
    END_IF;
    exPrev := Execute;
END_FUNCTION_BLOCK

// ---- FB_IotMqttReceive: poll for a pending publish ----
FUNCTION_BLOCK FB_IotMqttReceive
VAR_INPUT
    Execute : BOOL;
    ConnectionHdl : UDINT;
END_VAR
VAR_OUTPUT
    Done : BOOL;
    Message : BOOL;
    Error : BOOL;
    ErrorID : UDINT;
    Topic : STRING[127];
    Payload : STRING[255];
    PayloadLen : UDINT;
    QoS : UDINT;
    MessageId : UDINT;
    Retained : BOOL;
END_VAR
VAR
    ch : FB_Mqtt;
END_VAR
    Done := FALSE;
    Message := FALSE;
    Error := FALSE;
    ErrorID := 0;
    Retained := FALSE;
    IF Execute THEN
        ch.OP := 7;
        ch.HANDLE := ConnectionHdl;
        ch();
        IF ch.STATUS = 0 THEN
            Done := TRUE;
            Message := TRUE;
            Topic := ch.RXTOPIC;
            Payload := ch.RXPAYLOAD;
            PayloadLen := ch.RXPLEN;
            QoS := ch.RXQOS;
            MessageId := ch.RXMSGID;
            Retained := ch.RXRETAIN <> 0;
        ELSIF ch.STATUS = 1 THEN
            Done := TRUE;
        ELSE
            Error := TRUE;
            ErrorID := ch.ERRID;
        END_IF;
    END_IF;
END_FUNCTION_BLOCK

// ---- F_MqttTopicMatch: MQTT 3.1.1 topic-filter match ----
// '+' matches exactly one topic level, '#' matches the remaining
// levels (must be the last filter level).  Topic names and filters
// are bounded STRING[255]; matching is case-sensitive per spec.
// NOTE: no early RETURN (ST FUNCTION return semantics) — a match
// flag drives a single exit.
FUNCTION F_MqttTopicMatch : BOOL
VAR_INPUT
    Filter : STRING[255];
    Topic : STRING[255];
END_VAR
VAR
    f : STRING[255];
    t : STRING[255];
    fs : UDINT;
    ft : UDINT;
    fseg : STRING[255];
    tseg : STRING[255];
    fend : BOOL;
    match : BOOL;
END_VAR
    f := Filter;
    t := Topic;
    fend := FALSE;
    match := TRUE;
    WHILE NOT fend AND match DO
        IF LEN(f) = 0 THEN
            fend := TRUE;
        ELSE
            fs := FIND(f, '/');
            IF fs = 0 THEN
                fseg := f;
                f := '';
            ELSE
                fseg := LEFT(f, fs - 1);
                f := MID(f, LEN(f) - fs, fs + 1);
            END_IF;
            // '#' terminates the filter and matches the rest
            IF LEN(fseg) = 1 AND FIND(fseg, '#') = 1 THEN
                fend := TRUE;
                t := '';
            ELSE
                // consume the matching topic level
                IF LEN(t) = 0 THEN
                    tseg := '';
                ELSE
                    ft := FIND(t, '/');
                    IF ft = 0 THEN
                        tseg := t;
                        t := '';
                    ELSE
                        tseg := LEFT(t, ft - 1);
                        t := MID(t, LEN(t) - ft, ft + 1);
                    END_IF;
                END_IF;
                // '+' matches any single level
                IF LEN(fseg) = 1 AND FIND(fseg, '+') = 1 THEN
                    // matched; continue to next filter level
                ELSIF LEN(fseg) = 0 AND LEN(tseg) = 0 THEN
                    // empty==empty
                ELSIF LEN(fseg) > 0 AND LEN(tseg) > 0
                      AND LEN(fseg) = LEN(tseg) AND FIND(fseg, tseg) = 1 THEN
                    // literal level match
                ELSE
                    match := FALSE;
                END_IF;
            END_IF;
        END_IF;
    END_WHILE;
    // filter done: match only if topic is also exhausted
    F_MqttTopicMatch := match AND LEN(t) = 0;
END_FUNCTION

// ---- FB_IotMqttBackoff: Activate/DeactivateExponentialBackoff ----
// TwinCAT's ActivateExponentialBackoff(min,max) makes the client
// auto-reconnect with a doubling delay bounded by max; Deactivate
// stops it.  Enable=TRUE on the Execute edge activates with
// MinMs/MaxMs; Enable=FALSE deactivates.  Reconnects re-issue the
// original CONNECT (host/port/TLS/will); subscriptions are NOT
// restored — resubscribe after the connection returns.
FUNCTION_BLOCK FB_IotMqttBackoff
VAR_INPUT
    Execute : BOOL;
    ConnectionHdl : UDINT;
    MinMs : UDINT;
    MaxMs : UDINT;
    Enable : BOOL;
END_VAR
VAR_OUTPUT
    Done : BOOL;
    Error : BOOL;
    ErrorID : UDINT;
END_VAR
VAR
    ch : FB_Mqtt;
    exPrev : BOOL;
END_VAR
    Done := FALSE;
    Error := FALSE;
    ErrorID := 0;
    IF Execute AND NOT exPrev THEN
        ch.OP := 10;
        ch.HANDLE := ConnectionHdl;
        ch.BACKOFFMIN := MinMs;
        ch.BACKOFFMAX := MaxMs;
        IF Enable THEN ch.BACKOFFEN := 1; ELSE ch.BACKOFFEN := 0; END_IF;
        ch();
        IF ch.STATUS = 0 THEN
            Done := TRUE;
        ELSE
            Error := TRUE;
            ErrorID := ch.ERRID;
        END_IF;
    END_IF;
    exPrev := Execute;
END_FUNCTION_BLOCK

// ---- FB_IotMqttStatus: session status + broker-message age ----
// Level-triggered: while Execute is TRUE it polls the connection
// status each scan.  TimeSinceLastBrokerMsgMs is the
// GetTimeSinceLastBrokerMessage() equivalent — milliseconds since
// the last inbound broker message (PUBLISH delivery or connect;
// transport-level pings are not surfaced by the sync client).
FUNCTION_BLOCK FB_IotMqttStatus
VAR_INPUT
    Execute : BOOL;
    ConnectionHdl : UDINT;
END_VAR
VAR_OUTPUT
    Connected : BOOL;
    State : DINT;
    LastMsgId : UDINT;
    LastQos : UDINT;
    LastError : DINT;
    TimeSinceLastBrokerMsgMs : UDINT;
    Error : BOOL;
    ErrorID : UDINT;
END_VAR
VAR
    ch : FB_Mqtt;
END_VAR
    Connected := FALSE;
    Error := FALSE;
    ErrorID := 0;
    IF Execute THEN
        ch.OP := 3;
        ch.HANDLE := ConnectionHdl;
        ch();
        IF ch.STATUS = 0 THEN
            Connected := ch.STATE = 2;
            State := ch.STATE;
            LastMsgId := ch.LASTMSGID;
            LastError := ch.LASTERR;
            TimeSinceLastBrokerMsgMs := ch.LASTMSGSINCE;
        ELSE
            Error := TRUE;
            ErrorID := ch.ERRID;
        END_IF;
    END_IF;
END_FUNCTION_BLOCK

// ---- FB_IotMqttMessage: one queued MQTT message ----
// TwinCAT exposes GetTopic/GetPayload/CompareTopic methods; this
// dialect surfaces the same data as members.
FUNCTION_BLOCK FB_IotMqttMessage
VAR
    TOPIC : STRING[127];
    PAYLOAD : STRING[255];
    PAYLOADLEN : UDINT;
    QOS : UDINT;
    MSGID : UDINT;
    RETAINED : BOOL;
END_VAR
END_FUNCTION_BLOCK

// ---- FB_IotMqttMessageQueue: bounded FIFO of inbound messages ----
// TwinCAT's queue collects messages in the background and Dequeue
// transfers the oldest into an FB_IotMqttMessage.  This dialect has
// no REFERENCE TO inputs, so the popped message appears on the Msg*
// outputs instead.  Pump is level-triggered: each scan it drains up
// to 8 pending messages (bounded, watchdog-safe) into a 16-entry
// ring; DequeueReq/ResetReq are edge-triggered.
FUNCTION_BLOCK FB_IotMqttMessageQueue
VAR_INPUT
    Pump : BOOL;
    ConnectionHdl : UDINT;
    DequeueReq : BOOL;
    ResetReq : BOOL;
END_VAR
VAR_OUTPUT
    HasMessage : BOOL;
    Topic : STRING[127];
    Payload : STRING[255];
    PayloadLen : UDINT;
    QoS : UDINT;
    MessageId : UDINT;
    Retained : BOOL;
    Queued : UDINT;
    Error : BOOL;
    ErrorID : UDINT;
END_VAR
VAR
    head : UDINT;
    count : UDINT;
    qTopic : ARRAY[0..15] OF STRING[127];
    qPayload : ARRAY[0..15] OF STRING[255];
    qPayLen : ARRAY[0..15] OF UDINT;
    qQos : ARRAY[0..15] OF UDINT;
    qId : ARRAY[0..15] OF UDINT;
    qRet : ARRAY[0..15] OF BOOL;
    rx : FB_IotMqttReceive;
    slot : UDINT;
    dqPrev : BOOL;
    rsPrev : BOOL;
END_VAR
    HasMessage := FALSE;
    Error := FALSE;
    ErrorID := 0;
    IF Pump AND count < 16 THEN
        // one nonblocking receive per scan keeps the pump bounded
        rx.Execute := TRUE;
        rx.ConnectionHdl := ConnectionHdl;
        rx();
        rx.Execute := FALSE;
        IF rx.Message THEN
            slot := head + count;
            IF slot >= 16 THEN slot := slot - 16; END_IF;
            qTopic[slot] := rx.Topic;
            qPayload[slot] := rx.Payload;
            qPayLen[slot] := rx.PayloadLen;
            qQos[slot] := rx.QoS;
            qId[slot] := rx.MessageId;
            qRet[slot] := rx.Retained;
            count := count + 1;
        END_IF;
        IF rx.Error THEN
            Error := TRUE;
            ErrorID := rx.ErrorID;
        END_IF;
    END_IF;
    Queued := count;
    // dequeue: pop the oldest message into the Msg* outputs
    IF DequeueReq AND NOT dqPrev AND count > 0 THEN
        Topic := qTopic[head];
        Payload := qPayload[head];
        PayloadLen := qPayLen[head];
        QoS := qQos[head];
        MessageId := qId[head];
        Retained := qRet[head];
        HasMessage := TRUE;
        head := head + 1;
        IF head >= 16 THEN head := 0; END_IF;
        count := count - 1;
        Queued := count;
    END_IF;
    dqPrev := DequeueReq;
    // reset: drop every queued message
    IF ResetReq AND NOT rsPrev THEN
        head := 0;
        count := 0;
        Queued := 0;
    END_IF;
    rsPrev := ResetReq;
END_FUNCTION_BLOCK

// ---- FB_IotMqtt5Client: MQTT 5.0 CONNECT/CONNACK ----
// Same surface as FB_IotMqttClient plus the MQTT5 connect
// properties.  Publish/subscribe/unsubscribe reuse the existing
// FBs; the service picks the MQTT5 packet forms automatically for
// a v5 connection.
FUNCTION_BLOCK FB_IotMqtt5Client
VAR_INPUT
    Execute : BOOL;
    HostName : STRING[63];
    Port : UDINT;
    UserName : STRING[63];
    Password : STRING[127];
    ClientId : STRING[63];
    ConnectTimeoutMs : UDINT;
    MqttVersion : UDINT;      // 3|5
    Transport : UDINT;       // 0=auto 1=tcp 2=ssl 3=ws 4=wss
    CleanSession : BOOL;
    KeepAlive : UDINT;
    WillTopic : STRING[127];
    WillPayload : STRING[255];
    WillQoS : UDINT;
    WillRetain : BOOL;
    UseTls : BOOL;
    TlsInsecure : BOOL;
    TlsCaFile : STRING[127];
    TlsCertFile : STRING[127];
    TlsKeyFile : STRING[127];
    SessionExpiryS : UDINT;
    ReceiveMaximum : UDINT;
    TopicAliasMaximum : UDINT;
    RequestResponseInformation : BOOL;
    RequestProblemInformation : BOOL;
END_VAR
VAR_OUTPUT
    Done : BOOL;
    Busy : BOOL;
    Error : BOOL;
    ErrorID : UDINT;
    ConnectionHdl : UDINT;
END_VAR
VAR
    ch : FB_Mqtt;
    exPrev : BOOL;
END_VAR
    Done := FALSE;
    Error := FALSE;
    ErrorID := 0;
    IF Execute AND NOT exPrev THEN
        ch.OP := 1;
        ch.HOST := HostName;
        ch.PORT := Port;
        ch.USERNAME := UserName;
        ch.PASSWORD := Password;
        ch.CLIENTID := ClientId;
        ch.CONNECTMS := ConnectTimeoutMs;
        ch.MQTTVER := MqttVersion;
        ch.TRANSPORT := Transport;
        IF CleanSession THEN ch.CLEAN := 1; ELSE ch.CLEAN := 0; END_IF;
        ch.KEEPALIVE := KeepAlive;
        ch.WILLTOPIC := WillTopic;
        ch.WILLPAYLOAD := WillPayload;
        ch.WILLQOS := WillQoS;
        IF WillRetain THEN ch.WILLRETAIN := 1; ELSE ch.WILLRETAIN := 0; END_IF;
        IF UseTls THEN ch.USETLS := 1; ELSE ch.USETLS := 0; END_IF;
        IF TlsInsecure THEN ch.TLSINSECURE := 1; ELSE ch.TLSINSECURE := 0; END_IF;
        ch.TLSCAFILE := TlsCaFile;
        ch.TLSCERTFILE := TlsCertFile;
        ch.TLSKEYFILE := TlsKeyFile;
        ch.MQTTVER := 5;
        ch.M5SESSIONEXP := SessionExpiryS;
        ch.M5RECVMAX := ReceiveMaximum;
        ch.M5TOPICALIAS := TopicAliasMaximum;
        IF RequestResponseInformation THEN ch.M5REQRESP := 1; ELSE ch.M5REQRESP := 0; END_IF;
        IF RequestProblemInformation THEN ch.M5REQPROB := 1; ELSE ch.M5REQPROB := 0; END_IF;
        ch();
        IF ch.STATUS = 0 THEN
            Done := TRUE;
            ConnectionHdl := ch.HANDLE;
        ELSE
            Error := TRUE;
            ErrorID := ch.ERRID;
        END_IF;
    END_IF;
    exPrev := Execute;
    Busy := FALSE;
END_FUNCTION_BLOCK

// ---- FB_IotMqtt5Publish: MQTT5 PUBLISH with properties ----
// v5 connections only.  Property inputs map to
// TplcMqtt5PubProps; empty inputs leave the property absent.
// UserProperties is a "k1=v1;k2=v2" list.
FUNCTION_BLOCK FB_IotMqtt5Publish
VAR_INPUT
    Execute : BOOL;
    ConnectionHdl : UDINT;
    Topic : STRING[127];
    Payload : STRING[255];
    QoS : UDINT;
    RetainOn : BOOL;
    PayloadFormatUtf8 : BOOL;
    MessageExpiryS : UDINT;
    ContentType : STRING[127];
    ResponseTopic : STRING[127];
    CorrelationData : STRING[127];
    UserProperties : STRING[255];
END_VAR
VAR_OUTPUT
    Done : BOOL;
    Error : BOOL;
    ErrorID : UDINT;
END_VAR
VAR
    ch : FB_Mqtt;
    exPrev : BOOL;
END_VAR
    Done := FALSE;
    Error := FALSE;
    ErrorID := 0;
    IF Execute AND NOT exPrev THEN
        ch.OP := 11;
        ch.HANDLE := ConnectionHdl;
        ch.TOPIC := Topic;
        ch.PAYLOAD := Payload;
        ch.QOS := QoS;
        IF RetainOn THEN ch.FLG_RETAIN := 1; ELSE ch.FLG_RETAIN := 0; END_IF;
        IF PayloadFormatUtf8 THEN ch.M5PUBFMT := 1; ELSE ch.M5PUBFMT := 0; END_IF;
        ch.M5PUBEXPIRY := MessageExpiryS;
        ch.M5PUBCTYPE := ContentType;
        ch.M5PUBRTOPIC := ResponseTopic;
        ch.M5PUBCORR := CorrelationData;
        ch.M5PUBCORR_LEN := LEN(CorrelationData);
        ch.M5PUBUPROPS := UserProperties;
        ch();
        IF ch.STATUS = 0 THEN
            Done := TRUE;
        ELSE
            Error := TRUE;
            ErrorID := ch.ERRID;
        END_IF;
    END_IF;
    exPrev := Execute;
END_FUNCTION_BLOCK

// ---- FB_IotMqtt5Subscribe: MQTT5 SUBSCRIBE with properties ----
// v5 connections only.  NoLocal suppresses echoes of own
// publishes; RetainHandling: 0=always send retained, 1=new
// subscriptions only, 2=never.  SubscriptionId tags delivered
// messages; UserProperties is a "k1=v1;k2=v2" list.
FUNCTION_BLOCK FB_IotMqtt5Subscribe
VAR_INPUT
    Execute : BOOL;
    ConnectionHdl : UDINT;
    TopicFilter : STRING[127];
    QoS : UDINT;
    NoLocal : BOOL;
    RetainAsPublished : BOOL;
    RetainHandling : UDINT;
    SubscriptionId : UDINT;
    UserProperties : STRING[255];
END_VAR
VAR_OUTPUT
    Done : BOOL;
    Error : BOOL;
    ErrorID : UDINT;
END_VAR
VAR
    ch : FB_Mqtt;
    exPrev : BOOL;
END_VAR
    Done := FALSE;
    Error := FALSE;
    ErrorID := 0;
    IF Execute AND NOT exPrev THEN
        ch.OP := 12;
        ch.HANDLE := ConnectionHdl;
        ch.TOPIC := TopicFilter;
        ch.QOS := QoS;
        IF NoLocal THEN ch.M5SUBNOLOCAL := 1; ELSE ch.M5SUBNOLOCAL := 0; END_IF;
        IF RetainAsPublished THEN ch.M5SUBRAP := 1; ELSE ch.M5SUBRAP := 0; END_IF;
        ch.M5SUBRH := RetainHandling;
        ch.M5SUBSID := SubscriptionId;
        ch.M5SUBUPROPS := UserProperties;
        ch();
        IF ch.STATUS = 0 THEN
            Done := TRUE;
        ELSE
            Error := TRUE;
            ErrorID := ch.ERRID;
        END_IF;
    END_IF;
    exPrev := Execute;
END_FUNCTION_BLOCK

// ---- FB_IotMqtt5Receive: MQTT5 PUBLISH receive with properties ----
// v5 connections only.  Same poll semantics as FB_IotMqttReceive
// plus the PUBLISH property outputs: PayloadFormatUtf8,
// MessageExpiryS, SubscriptionId, ContentType, ResponseTopic,
// CorrelationData (STRING, binary-safe via LEN), UserProperties
// ("k=v;k=v" list).
FUNCTION_BLOCK FB_IotMqtt5Receive
VAR_INPUT
    Execute : BOOL;
    ConnectionHdl : UDINT;
END_VAR
VAR_OUTPUT
    Done : BOOL;
    Message : BOOL;
    Error : BOOL;
    ErrorID : UDINT;
    Topic : STRING[127];
    Payload : STRING[255];
    PayloadLen : UDINT;
    QoS : UDINT;
    MessageId : UDINT;
    Retained : BOOL;
    PayloadFormatUtf8 : BOOL;
    MessageExpiryS : UDINT;
    SubscriptionId : UDINT;
    ContentType : STRING[63];
    ResponseTopic : STRING[127];
    CorrelationData : STRING[127];
    CorrelationLen : UDINT;
    UserProperties : STRING[255];
END_VAR
VAR
    ch : FB_Mqtt;
END_VAR
    Done := FALSE;
    Message := FALSE;
    Error := FALSE;
    ErrorID := 0;
    Retained := FALSE;
    PayloadFormatUtf8 := FALSE;
    MessageExpiryS := 0;
    SubscriptionId := 0;
    CorrelationLen := 0;
    IF Execute THEN
        ch.OP := 13;
        ch.HANDLE := ConnectionHdl;
        ch();
        IF ch.STATUS = 0 THEN
            Done := TRUE;
            Message := TRUE;
            Topic := ch.RXTOPIC;
            Payload := ch.RXPAYLOAD;
            PayloadLen := ch.RXPLEN;
            QoS := ch.RXQOS;
            MessageId := ch.RXMSGID;
            Retained := ch.RXRETAIN <> 0;
            PayloadFormatUtf8 := ch.M5RXFMT <> 0;
            MessageExpiryS := ch.M5RXEXPIRY;
            SubscriptionId := ch.M5RXSUBID;
            ContentType := ch.M5RXCTYPE;
            ResponseTopic := ch.M5RXRTOPIC;
            CorrelationData := ch.M5RXCORR;
            CorrelationLen := ch.M5RXCORR_LEN;
            UserProperties := ch.M5RXUPROPS;
        ELSIF ch.STATUS = 1 THEN
            Done := TRUE;
        ELSE
            Error := TRUE;
            ErrorID := ch.ERRID;
        END_IF;
    END_IF;
END_FUNCTION_BLOCK

// ---- FB_IotMqtt5Message: one queued MQTT5 message ----
// TwinCAT's FB_IotMqtt5Message carries the PUBLISH property block
// alongside topic/payload; this dialect surfaces them as members.
FUNCTION_BLOCK FB_IotMqtt5Message
VAR
    TOPIC : STRING[127];
    PAYLOAD : STRING[255];
    PAYLOADLEN : UDINT;
    QOS : UDINT;
    MSGID : UDINT;
    RETAINED : BOOL;
    PAYLOADFORMATUTF8 : BOOL;
    MESSAGEEXPIRYS : UDINT;
    SUBSCRIPTIONID : UDINT;
    CONTENTTYPE : STRING[63];
    RESPONSETOPIC : STRING[127];
    CORRELATIONDATA : STRING[127];
    CORRELATIONLEN : UDINT;
    USERPROPERTIES : STRING[255];
END_VAR
END_FUNCTION_BLOCK

// ---- FB_IotMqtt5MessageQueue: bounded FIFO of inbound v5 msgs ----
// Same pump/dequeue model as FB_IotMqttMessageQueue but drains via
// FB_IotMqtt5Receive so queued entries keep the PUBLISH properties.
FUNCTION_BLOCK FB_IotMqtt5MessageQueue
VAR_INPUT
    Pump : BOOL;
    ConnectionHdl : UDINT;
    DequeueReq : BOOL;
    ResetReq : BOOL;
END_VAR
VAR_OUTPUT
    HasMessage : BOOL;
    Topic : STRING[127];
    Payload : STRING[255];
    PayloadLen : UDINT;
    QoS : UDINT;
    MessageId : UDINT;
    Retained : BOOL;
    PayloadFormatUtf8 : BOOL;
    MessageExpiryS : UDINT;
    SubscriptionId : UDINT;
    ContentType : STRING[63];
    ResponseTopic : STRING[127];
    CorrelationData : STRING[127];
    CorrelationLen : UDINT;
    UserProperties : STRING[255];
    Queued : UDINT;
    Error : BOOL;
    ErrorID : UDINT;
END_VAR
VAR
    head : UDINT;
    count : UDINT;
    qTopic : ARRAY[0..15] OF STRING[127];
    qPayload : ARRAY[0..15] OF STRING[255];
    qPayLen : ARRAY[0..15] OF UDINT;
    qQos : ARRAY[0..15] OF UDINT;
    qId : ARRAY[0..15] OF UDINT;
    qRet : ARRAY[0..15] OF BOOL;
    qFmt : ARRAY[0..15] OF BOOL;
    qExp : ARRAY[0..15] OF UDINT;
    qSub : ARRAY[0..15] OF UDINT;
    qCType : ARRAY[0..15] OF STRING[63];
    qRTopic : ARRAY[0..15] OF STRING[127];
    qCorr : ARRAY[0..15] OF STRING[127];
    qCorrLen : ARRAY[0..15] OF UDINT;
    qUProps : ARRAY[0..15] OF STRING[255];
    rx : FB_IotMqtt5Receive;
    slot : UDINT;
    dqPrev : BOOL;
    rsPrev : BOOL;
END_VAR
    HasMessage := FALSE;
    Error := FALSE;
    ErrorID := 0;
    IF Pump AND count < 16 THEN
        rx.Execute := TRUE;
        rx.ConnectionHdl := ConnectionHdl;
        rx();
        rx.Execute := FALSE;
        IF rx.Message THEN
            slot := head + count;
            IF slot >= 16 THEN slot := slot - 16; END_IF;
            qTopic[slot] := rx.Topic;
            qPayload[slot] := rx.Payload;
            qPayLen[slot] := rx.PayloadLen;
            qQos[slot] := rx.QoS;
            qId[slot] := rx.MessageId;
            qRet[slot] := rx.Retained;
            qFmt[slot] := rx.PayloadFormatUtf8;
            qExp[slot] := rx.MessageExpiryS;
            qSub[slot] := rx.SubscriptionId;
            qCType[slot] := rx.ContentType;
            qRTopic[slot] := rx.ResponseTopic;
            qCorr[slot] := rx.CorrelationData;
            qCorrLen[slot] := rx.CorrelationLen;
            qUProps[slot] := rx.UserProperties;
            count := count + 1;
        END_IF;
        IF rx.Error THEN
            Error := TRUE;
            ErrorID := rx.ErrorID;
        END_IF;
    END_IF;
    Queued := count;
    IF DequeueReq AND NOT dqPrev AND count > 0 THEN
        Topic := qTopic[head];
        Payload := qPayload[head];
        PayloadLen := qPayLen[head];
        QoS := qQos[head];
        MessageId := qId[head];
        Retained := qRet[head];
        PayloadFormatUtf8 := qFmt[head];
        MessageExpiryS := qExp[head];
        SubscriptionId := qSub[head];
        ContentType := qCType[head];
        ResponseTopic := qRTopic[head];
        CorrelationData := qCorr[head];
        CorrelationLen := qCorrLen[head];
        UserProperties := qUProps[head];
        HasMessage := TRUE;
        head := head + 1;
        IF head >= 16 THEN head := 0; END_IF;
        count := count - 1;
        Queued := count;
    END_IF;
    dqPrev := DequeueReq;
    IF ResetReq AND NOT rsPrev THEN
        head := 0;
        count := 0;
        Queued := 0;
    END_IF;
    rsPrev := ResetReq;
END_FUNCTION_BLOCK

// ---- FB_IotMqtt5RequestResponse: MQTT5 req/resp over the broker ----
// TwinCAT's Request/Response methods publish with ResponseTopic +
// CorrelationData properties and match the reply by correlation.
// This FB drives that flow as a bounded state machine: subscribe the
// response inbox once, publish the request, then poll
// FB_IotMqtt5Receive until a message whose Topic and CorrelationData
// match arrives (or TimeoutScans elapses -> Error).
FUNCTION_BLOCK FB_IotMqtt5RequestResponse
VAR_INPUT
    Execute : BOOL;
    ConnectionHdl : UDINT;
    RequestTopic : STRING[127];
    RequestPayload : STRING[255];
    QoS : UDINT;
    ResponseTopic : STRING[127];   // inbox to subscribe + advertise
    CorrelationData : STRING[127];
    TimeoutScans : UDINT;          // 0 = wait forever
END_VAR
VAR_OUTPUT
    Done : BOOL;
    Busy : BOOL;
    Error : BOOL;
    ErrorID : UDINT;
    ResponseTopicOut : STRING[127];
    ResponsePayload : STRING[255];
    ResponseQoS : UDINT;
    ResponseMessageId : UDINT;
END_VAR
VAR
    st : UDINT;
    waitN : UDINT;
    exPrev : BOOL;
    sub : FB_IotMqtt5Subscribe;
    pub : FB_IotMqtt5Publish;
    rx  : FB_IotMqtt5Receive;
END_VAR
    sub(); pub();
    Done := FALSE;
    Error := FALSE;
    ErrorID := 0;
    Busy := st <> 0;
    IF Execute AND NOT exPrev AND st = 0 THEN
        st := 1;
        waitN := 0;
    END_IF;
    exPrev := Execute;
    // st 1: subscribe the response inbox (once per request)
    IF st = 1 THEN
        sub.Execute := TRUE;
        sub.ConnectionHdl := ConnectionHdl;
        sub.TopicFilter := ResponseTopic;
        sub.QoS := 0;
        sub.NoLocal := FALSE;
        sub.RetainAsPublished := FALSE;
        sub.RetainHandling := 0;
        sub.SubscriptionId := 0;
        sub.UserProperties := '';
        st := 2;
    END_IF;
    IF st = 2 THEN
        IF sub.Done THEN
            sub.Execute := FALSE;
            pub.Execute := TRUE;
            pub.ConnectionHdl := ConnectionHdl;
            pub.Topic := RequestTopic;
            pub.Payload := RequestPayload;
            pub.QoS := QoS;
            pub.RetainOn := FALSE;
            pub.PayloadFormatUtf8 := FALSE;
            pub.MessageExpiryS := 0;
            pub.ContentType := '';
            pub.ResponseTopic := ResponseTopic;
            pub.CorrelationData := CorrelationData;
            pub.UserProperties := '';
            st := 3;
        END_IF;
        IF sub.Error THEN
            Error := TRUE; ErrorID := sub.ErrorID; st := 0;
        END_IF;
    END_IF;
    IF st = 3 THEN
        IF pub.Done THEN
            pub.Execute := FALSE;
            st := 4;
        END_IF;
        IF pub.Error THEN
            Error := TRUE; ErrorID := pub.ErrorID; st := 0;
        END_IF;
    END_IF;
    // st 4: poll for the correlated response
    IF st = 4 THEN
        rx.Execute := TRUE;
        rx.ConnectionHdl := ConnectionHdl;
        rx();
        rx.Execute := FALSE;
        IF rx.Message THEN
            IF rx.Topic = ResponseTopic
               AND rx.CorrelationData = CorrelationData THEN
                ResponseTopicOut := rx.Topic;
                ResponsePayload := rx.Payload;
                ResponseQoS := rx.QoS;
                ResponseMessageId := rx.MessageId;
                Done := TRUE;
                st := 0;
            END_IF;
        END_IF;
        IF rx.Error THEN
            Error := TRUE; ErrorID := rx.ErrorID; st := 0;
        END_IF;
        waitN := waitN + 1;
        IF TimeoutScans > 0 AND waitN >= TimeoutScans THEN
            Error := TRUE; ErrorID := 90; st := 0;
        END_IF;
    END_IF;
END_FUNCTION_BLOCK

// ---- MQTT5 property containers (Tc3_IotBase §5.1.2.9) ----
// TwinCAT passes these FBs by reference into the client methods.
// This dialect has no REFERENCE TO parameters, so the publish and
// subscribe FBs take the same fields as direct inputs; these
// containers give user code a named place to stage property values
// before copying them onto FB_IotMqtt5Publish/Subscribe inputs.

// FB_IotMqtt5ConnAckProperties: broker properties received in the
// CONNACK (session expiry, receive maximum, topic alias maximum,
// reason string, user properties).
FUNCTION_BLOCK FB_IotMqtt5ConnAckProperties
VAR
    SessionExpiryInterval : UDINT;
    ReceiveMaximum : UDINT;
    TopicAliasMaximum : UDINT;
    ReasonString : STRING[127];
    UserProperties : STRING[255];
END_VAR
END_FUNCTION_BLOCK

// FB_IotMqtt5DisconnectProperties: properties received in the
// broker's DISCONNECT (reason code, reason string, session expiry,
// user properties).
FUNCTION_BLOCK FB_IotMqtt5DisconnectProperties
VAR
    ReasonCode : UDINT;
    ReasonString : STRING[127];
    SessionExpiryInterval : UDINT;
    UserProperties : STRING[255];
END_VAR
END_FUNCTION_BLOCK

// FB_IotMqtt5PublishProperties: properties attached to an outgoing
// PUBLISH (payload format, message expiry, content type, response
// topic, correlation data, user properties).
FUNCTION_BLOCK FB_IotMqtt5PublishProperties
VAR
    PayloadFormatIndicator : BOOL;
    MessageExpiryInterval : UDINT;
    ContentType : STRING[63];
    ResponseTopic : STRING[127];
    CorrelationData : STRING[127];
    CorrelationDataLen : UDINT;
    UserProperties : STRING[255];
END_VAR
END_FUNCTION_BLOCK

// FB_IotMqtt5SubscribeProperties: properties attached to a
// SUBSCRIBE (no-local, retain-as-published, retain handling,
// subscription identifier, user properties).
FUNCTION_BLOCK FB_IotMqtt5SubscribeProperties
VAR
    NoLocal : BOOL;
    RetainAsPublished : BOOL;
    RetainHandling : UDINT;
    SubscriptionIdentifier : UDINT;
    UserProperties : STRING[255];
END_VAR
END_FUNCTION_BLOCK

// FB_IotMqtt5UnsubscribeProperties: properties attached to an
// UNSUBSCRIBE (user properties only per MQTT5).
FUNCTION_BLOCK FB_IotMqtt5UnsubscribeProperties
VAR
    UserProperties : STRING[255];
END_VAR
END_FUNCTION_BLOCK

// FB_IotMqtt5UserProperties: bounded key/value list used to build
// the "k=v;k=v" encoding consumed by the property inputs above.
// AddReq appends one pair per call; the encoded list is on
// Encoded.  8 pairs max.
FUNCTION_BLOCK FB_IotMqtt5UserProperties
VAR_INPUT
    AddReq : BOOL;
    PropKey : STRING[63];
    PropValue : STRING[127];
    ClearReq : BOOL;
END_VAR
VAR_OUTPUT
    Count : UDINT;
    Encoded : STRING[255];
END_VAR
VAR
    n : UDINT;
    i : UDINT;
    keys : ARRAY[0..7] OF STRING[63];
    vals : ARRAY[0..7] OF STRING[127];
    addPrev : BOOL;
    clrPrev : BOOL;
END_VAR
    Count := n;
    Encoded := '';
    IF AddReq AND NOT addPrev AND n < 8 AND PropKey <> '' THEN
        keys[n] := PropKey;
        vals[n] := PropValue;
        n := n + 1;
    END_IF;
    addPrev := AddReq;
    IF ClearReq AND NOT clrPrev THEN
        n := 0;
    END_IF;
    clrPrev := ClearReq;
    // rebuild the k=v;k=v encoding
    IF n > 0 THEN
        Encoded := CONCAT(keys[0], CONCAT('=', vals[0]));
        FOR i := 1 TO n - 1 DO
            Encoded := CONCAT(Encoded, CONCAT(';',
                CONCAT(keys[i], CONCAT('=', vals[i]))));
        END_FOR;
    END_IF;
    Count := n;
END_FUNCTION_BLOCK

(* ---- tc2_ncfifoaxes.st ---- *)
// tc2_ncfifoaxes.st — Tc2_NcFifoAxes: FiFoAxes synchronous numeric
// setpoint FIFO channels (8 APIs) over the tplc-fifo service /
// FB_Fifo builtin.
//
// A FIFO channel queues rows of LREAL target positions (one column
// per integrated axis, group position = column) and emits one row
// per drive-clock tick as DS402 0x607A CSP targets. This is the
// numeric FiFoAxes surface; it is NOT the NC channel's G-code block
// queue (FB_ItpFiFoWrite / nc.fifo in tc2_nci.st).
//
// Flattening vs the TwinCAT signatures:
//   iChannelId    -> iChannelId (UDINT, 0..TPLC_FIFO_CHAN_MAX-1)
//   iAxisId       -> axis handle (UDINT; the same handle space as
//                    AXIS_REF / FB_MotionAxis, slave = handle-1 on
//                    Tether IO)
//   iGroupPosition-> 1-based in TwinCAT; mapped to the 0-based wire
//                    column internally
//   AdrDataArray  -> AdrDataArray : ARRAY[0..255] OF LREAL (flattened
//                    POINTER TO LREAL; the caller fills the wrapper's
//                    array, iRowsToWrite bounds the valid prefix,
//                    max 31 rows per call — chunk larger streams)
//   tTimeout      -> accepted, ignored (service calls are synchronous)
//   outputs       -> bBusy / bError / nErrorId plus domain outputs;
//                    bBusy pulses TRUE only during the Execute edge
// Channel state is visible on the internal FB_Fifo instance fields
// (STATE/QLEN/SEQ/NAXES/MAXROWS) for callers that need polling.

// ---- FiFoGetDimension: axes + capacity of a channel ----
FUNCTION_BLOCK FiFoGetDimension
VAR_INPUT
    iChannelId : UDINT;
    bExecute : BOOL;
    tTimeout : TIME;
END_VAR
VAR_OUTPUT
    bBusy : BOOL;
    bError : BOOL;
    nErrorId : UDINT;
    iAxes : UDINT;
    iMaxRows : UDINT;
END_VAR
VAR
    ch : FB_Fifo;
    exPrev : BOOL;
END_VAR
    bBusy := FALSE;
    bError := FALSE;
    nErrorId := 0;
    IF bExecute AND NOT exPrev THEN
        bBusy := TRUE;
        ch.OP := 8;
        ch.CHAN := iChannelId;
        ch();
        IF ch.STATUS = 0 THEN
            iAxes := ch.NAXES;
            iMaxRows := ch.MAXROWS;
        ELSE
            bError := TRUE;
            nErrorId := ch.ERRID;
        END_IF;
    END_IF;
    exPrev := bExecute;
END_FUNCTION_BLOCK

// ---- FiFoGroupIntegrate: add an axis to the channel ----
FUNCTION_BLOCK FiFoGroupIntegrate
VAR_INPUT
    iChannelId : UDINT;
    iAxisId : UDINT;
    iGroupPosition : UDINT;
    bExecute : BOOL;
    tTimeout : TIME;
END_VAR
VAR_OUTPUT
    bBusy : BOOL;
    bError : BOOL;
    nErrorId : UDINT;
END_VAR
VAR
    ch : FB_Fifo;
    exPrev : BOOL;
END_VAR
    bBusy := FALSE;
    bError := FALSE;
    nErrorId := 0;
    IF bExecute AND NOT exPrev THEN
        bBusy := TRUE;
        ch.OP := 1;
        ch.CHAN := iChannelId;
        /* TwinCAT group positions are 1-based; the wire column is
           0-based. */
        ch.AUX := iAxisId OR ((iGroupPosition - 1) * 65536);
        ch();
        IF ch.STATUS <> 0 THEN
            bError := TRUE;
            nErrorId := ch.ERRID;
        END_IF;
    END_IF;
    exPrev := bExecute;
END_FUNCTION_BLOCK

// ---- FiFoGroupDisintegrate: clear axes + queued rows ----
FUNCTION_BLOCK FiFoGroupDisintegrate
VAR_INPUT
    iChannelId : UDINT;
    bExecute : BOOL;
    tTimeout : TIME;
END_VAR
VAR_OUTPUT
    bBusy : BOOL;
    bError : BOOL;
    nErrorId : UDINT;
END_VAR
VAR
    ch : FB_Fifo;
    exPrev : BOOL;
END_VAR
    bBusy := FALSE;
    bError := FALSE;
    nErrorId := 0;
    IF bExecute AND NOT exPrev THEN
        bBusy := TRUE;
        ch.OP := 2;
        ch.CHAN := iChannelId;
        ch();
        IF ch.STATUS <> 0 THEN
            bError := TRUE;
            nErrorId := ch.ERRID;
        END_IF;
    END_IF;
    exPrev := bExecute;
END_FUNCTION_BLOCK

// ---- FiFoWrite / FiFoOverwrite shared row pump ----
// Both copy caller rows into the FB_Fifo ROWS staging buffer in
// chunks of 32 rows (256 LREAL) and issue OP3 (append) / OP4
// (replace queue first) per chunk.
FUNCTION_BLOCK FiFoWritePump
VAR_INPUT
    iChannelId : UDINT;
    AdrDataArray : ARRAY[0..255] OF LREAL;
    iRowsToWrite : UDINT;
    bOverwrite : BOOL;
    bExecute : BOOL;
    tTimeout : TIME;
END_VAR
VAR_OUTPUT
    bBusy : BOOL;
    bError : BOOL;
    nErrorId : UDINT;
END_VAR
VAR
    ch : FB_Fifo;
    exPrev : BOOL;
    i : UDINT;
    r : UDINT;
    n : UDINT;
    base : UDINT;
END_VAR
    bBusy := FALSE;
    bError := FALSE;
    nErrorId := 0;
    IF bExecute AND NOT exPrev THEN
        bBusy := TRUE;
        i := 0;
        WHILE i < iRowsToWrite AND NOT bError DO
            n := iRowsToWrite - i;
            IF n > 32 THEN n := 32; END_IF;
            ch.OP := 3;
            IF bOverwrite THEN ch.OP := 4; END_IF;
            ch.CHAN := iChannelId;
            ch.NROWS := n;
            base := i * 8;
            FOR r := 0 TO 255 DO
                ch.ROWS[r] := 0.0;
            END_FOR;
            FOR r := 0 TO n * 8 - 1 DO
                ch.ROWS[r] := AdrDataArray[base + r];
            END_FOR;
            ch();
            IF ch.STATUS <> 0 THEN
                bError := TRUE;
                nErrorId := ch.ERRID;
            END_IF;
            i := i + n;
        END_WHILE;
    END_IF;
    exPrev := bExecute;
END_FUNCTION_BLOCK

FUNCTION_BLOCK FiFoWrite
VAR_INPUT
    iChannelId : UDINT;
    AdrDataArray : ARRAY[0..255] OF LREAL;
    iRowsToWrite : UDINT;
    bExecute : BOOL;
    tTimeout : TIME;
END_VAR
VAR_OUTPUT
    bBusy : BOOL;
    bError : BOOL;
    nErrorId : UDINT;
END_VAR
VAR
    pump : FiFoWritePump;
END_VAR
    pump.iChannelId := iChannelId;
    pump.AdrDataArray := AdrDataArray;
    pump.iRowsToWrite := iRowsToWrite;
    pump.bOverwrite := FALSE;
    pump.bExecute := bExecute;
    pump.tTimeout := tTimeout;
    pump();
    bBusy := pump.bBusy;
    bError := pump.bError;
    nErrorId := pump.nErrorId;
END_FUNCTION_BLOCK

FUNCTION_BLOCK FiFoOverwrite
VAR_INPUT
    iChannelId : UDINT;
    AdrDataArray : ARRAY[0..255] OF LREAL;
    iRowsToWrite : UDINT;
    bExecute : BOOL;
    tTimeout : TIME;
END_VAR
VAR_OUTPUT
    bBusy : BOOL;
    bError : BOOL;
    nErrorId : UDINT;
END_VAR
VAR
    pump : FiFoWritePump;
END_VAR
    pump.iChannelId := iChannelId;
    pump.AdrDataArray := AdrDataArray;
    pump.iRowsToWrite := iRowsToWrite;
    pump.bOverwrite := TRUE;
    pump.bExecute := bExecute;
    pump.tTimeout := tTimeout;
    pump();
    bBusy := pump.bBusy;
    bError := pump.bError;
    nErrorId := pump.nErrorId;
END_FUNCTION_BLOCK

// ---- FiFoStart: begin streaming queued rows ----
FUNCTION_BLOCK FiFoStart
VAR_INPUT
    iChannelId : UDINT;
    bExecute : BOOL;
    tTimeout : TIME;
END_VAR
VAR_OUTPUT
    bBusy : BOOL;
    bError : BOOL;
    nErrorId : UDINT;
END_VAR
VAR
    ch : FB_Fifo;
    exPrev : BOOL;
END_VAR
    bBusy := FALSE;
    bError := FALSE;
    nErrorId := 0;
    IF bExecute AND NOT exPrev THEN
        bBusy := TRUE;
        ch.OP := 5;
        ch.CHAN := iChannelId;
        ch.AUX := 1;
        ch();
        IF ch.STATUS <> 0 THEN
            bError := TRUE;
            nErrorId := ch.ERRID;
        END_IF;
    END_IF;
    exPrev := bExecute;
END_FUNCTION_BLOCK

// ---- FiFoStop: halt the channel (queued rows kept) ----
FUNCTION_BLOCK FiFoStop
VAR_INPUT
    iChannelId : UDINT;
    bExecute : BOOL;
    tTimeout : TIME;
END_VAR
VAR_OUTPUT
    bBusy : BOOL;
    bError : BOOL;
    nErrorId : UDINT;
END_VAR
VAR
    ch : FB_Fifo;
    exPrev : BOOL;
END_VAR
    bBusy := FALSE;
    bError := FALSE;
    nErrorId := 0;
    IF bExecute AND NOT exPrev THEN
        bBusy := TRUE;
        ch.OP := 5;
        ch.CHAN := iChannelId;
        ch.AUX := 2;
        ch();
        IF ch.STATUS <> 0 THEN
            bError := TRUE;
            nErrorId := ch.ERRID;
        END_IF;
    END_IF;
    exPrev := bExecute;
END_FUNCTION_BLOCK

// ---- FiFoSetChannelOverride: override percent (recorded) ----
FUNCTION_BLOCK FiFoSetChannelOverride
VAR_INPUT
    iChannelId : UDINT;
    iOverride : UDINT;
    bExecute : BOOL;
    tTimeout : TIME;
END_VAR
VAR_OUTPUT
    bBusy : BOOL;
    bError : BOOL;
    nErrorId : UDINT;
END_VAR
VAR
    ch : FB_Fifo;
    exPrev : BOOL;
END_VAR
    bBusy := FALSE;
    bError := FALSE;
    nErrorId := 0;
    IF bExecute AND NOT exPrev THEN
        bBusy := TRUE;
        ch.OP := 7;
        ch.CHAN := iChannelId;
        ch.VAL := UDINT_TO_LREAL(iOverride);
        ch();
        IF ch.STATUS <> 0 THEN
            bError := TRUE;
            nErrorId := ch.ERRID;
        END_IF;
    END_IF;
    exPrev := bExecute;
END_FUNCTION_BLOCK

FUNCTION F_GetVersionTcFifoAxes : STRING[32]
    F_GetVersionTcFifoAxes := 'Tc2_NcFifoAxes 1.0';
END_FUNCTION
